	IF stCmdModesStates.stStates.Active THEN
		stCmdModesStates.stStates.Active := FALSE;
		gpCh[nChanIdx]^.channel_mc_control.mode_and_state.command_w.to_mode := HLI_IMCM_AUTOMATIC_MODE;
		gpCh[nChanIdx]^.channel_mc_control.mode_and_state.command_w.to_state := HLI_IMCM_PROCESS_ACTIVE;		
		pString := ADR(gpCh[nChanIdx]^.channel_mc_control.mode_and_state.command_w.parameter);			
		pString^ := ProgramName;				
		gpCh[nChanIdx]^.channel_mc_control.mode_and_state.command_semaphor_rw  := TRUE;		
	END_IF
	
	IF stCmdModesStates.stStates.Hold THEN
		stCmdModesStates.stStates.Hold:= FALSE;
		gpCh[nChanIdx]^.channel_mc_control.mode_and_state.command_w.to_mode:= HLI_IMCM_AUTOMATIC_MODE;
		gpCh[nChanIdx]^.channel_mc_control.mode_and_state.command_w.to_state := HLI_IMCM_PROCESS_HOLD;		
		gpCh[nChanIdx]^.channel_mc_control.mode_and_state.command_semaphor_rw  := TRUE;
	END_IF
	
	IF stCmdModesStates.stStates.Reset THEN
		stCmdModesStates.stStates.Reset := FALSE;
		gpCh[nChanIdx]^.channel_mc_control.mode_and_state.command_w.to_mode := HLI_IMCM_AUTOMATIC_MODE;
		gpCh[nChanIdx]^.channel_mc_control.mode_and_state.command_w.to_state:= HLI_IMCM_PROCESS_RESETTING;		
		gpCh[nChanIdx]^.channel_mc_control.mode_and_state.command_semaphor_rw  := TRUE;		
	END_IF
	
	HLI3_ChannelModeAuto := TRUE;
ELSE
	HLI3_ChannelModeAuto := FALSE;
END_IF

END_FUNCTION

// CNC/2 OperationMode/HLI3_ChannelModeManual
FUNCTION HLI3_ChannelModeManual : BOOL
VAR_INPUT	
	nChanIdx: INT;	
END_VAR

VAR_IN_OUT
	stCmdModesStates    : ST_CNCCmdModesStates;	
END_VAR

VAR
	pString: POINTER TO STRING;
END_VAR

(* ========================================================= *)
(*    FUN: HLI_ChannelModeManual                             *)
(* --------------------------------------------------------- *)
(*   Desc: switch channel to Manual mode / xxx               *)
(*   Author: MK, MiB, TV, RCH                                *)
(*   Date: 03.03.2017                                        *)
(*   Rev.: 1.5                                               *)
(* ========================================================= *)

IF (NOT  gpCh[nChanIdx]^.channel_mc_control.mode_and_state.command_semaphor_rw) THEN    (* only if semaphor is FALSE...... *)
	IF stCmdModesStates.stStates.Selected THEN
		stCmdModesStates.stStates.Selected := FALSE;
		gpCh[nChanIdx]^.channel_mc_control.mode_and_state.command_w.to_mode := HLI_IMCM_MANUAL_MODE;
		gpCh[nChanIdx]^.channel_mc_control.mode_and_state.command_w.to_state := HLI_IMCM_PROCESS_SELECTED;		
		pString := ADR(gpCh[nChanIdx]^.channel_mc_control.mode_and_state.command_w.parameter);			
		pString^ := '';	
		gpCh[nChanIdx]^.channel_mc_control.mode_and_state.command_semaphor_rw := TRUE;		
	END_IF
	
	IF stCmdModesStates.stStates.Ready THEN
		stCmdModesStates.stStates.Ready := FALSE;
		gpCh[nChanIdx]^.channel_mc_control.mode_and_state.command_w.to_mode := HLI_IMCM_MANUAL_MODE;
		gpCh[nChanIdx]^.channel_mc_control.mode_and_state.command_w.to_state := HLI_IMCM_PROCESS_READY;		
		pString := ADR(gpCh[nChanIdx]^.channel_mc_control.mode_and_state.command_w.parameter);			
		pString^ := '';
		gpCh[nChanIdx]^.channel_mc_control.mode_and_state.command_semaphor_rw := TRUE;		
	END_IF
	
	IF stCmdModesStates.stStates.Active THEN
		stCmdModesStates.stStates.Active := FALSE;
		gpCh[nChanIdx]^.channel_mc_control.mode_and_state.command_w.to_mode := HLI_IMCM_MANUAL_MODE;
		gpCh[nChanIdx]^.channel_mc_control.mode_and_state.command_w.to_state := HLI_IMCM_PROCESS_ACTIVE;		
		pString := ADR(gpCh[nChanIdx]^.channel_mc_control.mode_and_state.command_w.parameter);			
		pString^ := '';						
		gpCh[nChanIdx]^.channel_mc_control.mode_and_state.command_semaphor_rw := TRUE;	
	END_IF
	
	IF stCmdModesStates.stStates.Hold THEN
		stCmdModesStates.stStates.Hold := FALSE;
		gpCh[nChanIdx]^.channel_mc_control.mode_and_state.command_w.to_mode := HLI_IMCM_MANUAL_MODE;
		gpCh[nChanIdx]^.channel_mc_control.mode_and_state.command_w.to_state := HLI_IMCM_PROCESS_HOLD;		
		gpCh[nChanIdx]^.channel_mc_control.mode_and_state.command_semaphor_rw := TRUE;		
	END_IF
	
	IF stCmdModesStates.stStates.Reset THEN
		stCmdModesStates.stStates.Reset := FALSE;
		gpCh[nChanIdx]^.channel_mc_control.mode_and_state.command_w.to_mode:= HLI_IMCM_MANUAL_MODE;
		gpCh[nChanIdx]^.channel_mc_control.mode_and_state.command_w.to_state := HLI_IMCM_PROCESS_RESETTING;		
		gpCh[nChanIdx]^.channel_mc_control.mode_and_state.command_semaphor_rw:= TRUE;		
	END_IF

	HLI3_ChannelModeManual := TRUE;
ELSE
	HLI3_ChannelModeManual := FALSE;
END_IF

END_FUNCTION

// CNC/2 OperationMode/HLI3_ChannelModeMDI
FUNCTION HLI3_ChannelModeMDI : BOOL
VAR_INPUT	
	nChanIdx: INT;	
	/// pointer to the MDI program string 
	pMDIString: POINTER TO STRING(HLI_IMCM_MODE_STATE_PARAM_STRL);
END_VAR

VAR_IN_OUT
	stCmdModesStates    : ST_CNCCmdModesStates;	
END_VAR
VAR
	pString: POINTER TO STRING(HLI_IMCM_MODE_STATE_PARAM_STRL);
END_VAR

(* ========================================================= *)
(*    FUN: HLI_ChannelModeMDI                                *)
(* --------------------------------------------------------- *)
(*   Desc: switch channel to MDI mode / xxx                  *)
(*   Author: MK, TV, MiB, Rch                                *)
(*   Date: 18.07.2002                                        *)
(*   Last: 03.03.2017                      				     *)
(*   Rev.: 1.7                                               *)
(* ========================================================= *)

IF (NOT gpCh[nChanIdx]^.channel_mc_control.mode_and_state.command_semaphor_rw) THEN  (* only if semaphor is FALSE...... *)

	IF stCmdModesStates.stStates.Selected THEN
		stCmdModesStates.stStates.Selected := FALSE;
		gpCh[nChanIdx]^.channel_mc_control.mode_and_state.command_w.to_mode := HLI_IMCM_MDI_MODE;
		gpCh[nChanIdx]^.channel_mc_control.mode_and_state.command_w.to_state := HLI_IMCM_PROCESS_SELECTED;
		pString := ADR(gpCh[nChanIdx]^.channel_mc_control.mode_and_state.command_w.parameter);					
		pString^ := pMDIString^;
		gpCh[nChanIdx]^.channel_mc_control.mode_and_state.command_semaphor_rw := TRUE;		
	END_IF
	
	IF stCmdModesStates.stStates.Ready THEN
		stCmdModesStates.stStates.Ready := FALSE;
		gpCh[nChanIdx]^.channel_mc_control.mode_and_state.command_w.to_mode:= HLI_IMCM_MDI_MODE;
		gpCh[nChanIdx]^.channel_mc_control.mode_and_state.command_w.to_state := HLI_IMCM_PROCESS_READY;		
		gpCh[nChanIdx]^.channel_mc_control.mode_and_state.command_semaphor_rw := TRUE;		
	END_IF
	
	IF stCmdModesStates.stStates.Active THEN
		stCmdModesStates.stStates.Active := FALSE;
		gpCh[nChanIdx]^.channel_mc_control.mode_and_state.command_w.to_mode := HLI_IMCM_MDI_MODE;
		gpCh[nChanIdx]^.channel_mc_control.mode_and_state.command_w.to_state := HLI_IMCM_PROCESS_ACTIVE;
		pString := ADR(gpCh[nChanIdx]^.channel_mc_control.mode_and_state.command_w.parameter);					
		pString^ := pMDIString^;
		gpCh[nChanIdx]^.channel_mc_control.mode_and_state.command_semaphor_rw := TRUE;		
	END_IF
	
	IF stCmdModesStates.stStates.Hold THEN
		stCmdModesStates.stStates.Hold := FALSE;
		gpCh[nChanIdx]^.channel_mc_control.mode_and_state.command_w.to_mode := HLI_IMCM_MDI_MODE;
		gpCh[nChanIdx]^.channel_mc_control.mode_and_state.command_w.to_state:= HLI_IMCM_PROCESS_HOLD;		
		gpCh[nChanIdx]^.channel_mc_control.mode_and_state.command_semaphor_rw := TRUE;		
	END_IF
	
	IF stCmdModesStates.stStates.Reset THEN
		stCmdModesStates.stStates.Reset := FALSE;
		gpCh[nChanIdx]^.channel_mc_control.mode_and_state.command_w.to_mode := HLI_IMCM_MDI_MODE;
		gpCh[nChanIdx]^.channel_mc_control.mode_and_state.command_w.to_state := HLI_IMCM_PROCESS_RESETTING;		
		gpCh[nChanIdx]^.channel_mc_control.mode_and_state.command_semaphor_rw := TRUE;		
	END_IF
	HLI3_ChannelModeMDI := TRUE;	
ELSE
	HLI3_ChannelModeMDI := FALSE;
END_IF

END_FUNCTION

// CNC/2 OperationMode/HLI3_ChannelModeReference
FUNCTION HLI3_ChannelModeReference : BOOL
VAR_INPUT	
	nChanIdx: INT;	
	/// the referencing string 
	sRefPosString: STRING(HLI_IMCM_MODE_STATE_PARAM_STRL);	
END_VAR

VAR_IN_OUT
	stCmdModesStates    : ST_CNCCmdModesStates;	
END_VAR

VAR
	pString: POINTER TO STRING(HLI_IMCM_MODE_STATE_PARAM_STRL);
END_VAR

(* ========================================================= *)
(*    FUN: HLI_ChannelModeReference                          *)
(* --------------------------------------------------------- *)
(*   Desc: switch channel to Reference mode / xxx            *)
(*   Author: MK, MiB, TV                                     *)
(*   Date: 03.03.2017                                        *)
(*   Rev.: 1.5                                               *)
(* ========================================================= *)


(************************************************************
	RefPosString:
	Element: parameter ( ASCII char set, Länge:256 Zeichen)

	Vorgabe zur Parametrierung der Referenzpunktfahrt.

	Ist dieser STRING leer, so wird defaultmäßig das
	Automatikprogramm "rpf.nc" angewählt.

	Ansonsten kann durch explizite Angabe der Achsen und
	Zeitpunkt im Format "G74
	<Achsbezeichner_1><Zeitpunkt_1> ...
	<Achsbezeichner_n><Zeitpunkt_n>"
	eine individuelle Referenzpunktfahrt vorgegeben werden.
*************************************************************)

IF (NOT gpCh[nChanIdx]^.channel_mc_control.mode_and_state.command_semaphor_rw) THEN  (* only if semaphor is FALSE...... *)
	IF stCmdModesStates.stStates.Selected THEN
		stCmdModesStates.stStates.Selected := FALSE;
		gpCh[nChanIdx]^.channel_mc_control.mode_and_state.command_w.to_mode := HLI_IMCM_REFERENCE_MODE;
		gpCh[nChanIdx]^.channel_mc_control.mode_and_state.command_w.to_state := HLI_IMCM_PROCESS_SELECTED;		
		gpCh[nChanIdx]^.channel_mc_control.mode_and_state.command_semaphor_rw := TRUE;	
	END_IF
	
	IF stCmdModesStates.stStates.Ready THEN
		stCmdModesStates.stStates.Ready := FALSE;
		gpCh[nChanIdx]^.channel_mc_control.mode_and_state.command_w.to_mode := HLI_IMCM_REFERENCE_MODE;
		gpCh[nChanIdx]^.channel_mc_control.mode_and_state.command_w.to_state := HLI_IMCM_PROCESS_READY;		
		pString := ADR(gpCh[nChanIdx]^.channel_mc_control.mode_and_state.command_w.parameter);	
		gpCh[nChanIdx]^.channel_mc_control.mode_and_state.command_semaphor_rw := TRUE;		
	END_IF
	
	IF stCmdModesStates.stStates.Active THEN
		stCmdModesStates.stStates.Active := FALSE;
		gpCh[nChanIdx]^.channel_mc_control.mode_and_state.command_w.to_mode := HLI_IMCM_REFERENCE_MODE;
		gpCh[nChanIdx]^.channel_mc_control.mode_and_state.command_w.to_state := HLI_IMCM_PROCESS_ACTIVE;		
		pString := ADR(gpCh[nChanIdx]^.channel_mc_control.mode_and_state.command_w.parameter);	
		pString^ := sRefPosString;
		gpCh[nChanIdx]^.channel_mc_control.mode_and_state.command_semaphor_rw:= TRUE;		
	END_IF
	
	IF stCmdModesStates.stStates.Hold THEN
		stCmdModesStates.stStates.Hold := FALSE;
		gpCh[nChanIdx]^.channel_mc_control.mode_and_state.command_w.to_mode := HLI_IMCM_REFERENCE_MODE;
		gpCh[nChanIdx]^.channel_mc_control.mode_and_state.command_w.to_state := HLI_IMCM_PROCESS_HOLD;		
		gpCh[nChanIdx]^.channel_mc_control.mode_and_state.command_semaphor_rw := TRUE;		
	END_IF
	
	IF stCmdModesStates.stStates.Reset THEN
		stCmdModesStates.stStates.Reset := FALSE;
		gpCh[nChanIdx]^.channel_mc_control.mode_and_state.command_w.to_mode:= HLI_IMCM_REFERENCE_MODE;
		gpCh[nChanIdx]^.channel_mc_control.mode_and_state.command_w.to_state := HLI_IMCM_PROCESS_RESETTING;		
		gpCh[nChanIdx]^.channel_mc_control.mode_and_state.command_semaphor_rw := TRUE;		
	END_IF

	HLI3_ChannelModeReference := TRUE;
ELSE
	HLI3_ChannelModeReference := FALSE;
END_IF

END_FUNCTION

// CNC/2 OperationMode/HLI3_ChannelModeStandby
FUNCTION HLI3_ChannelModeStandby : BOOL
VAR_INPUT	 
	nChanIdx: INT;
	ProgramName: STRING(HLI_IMCM_MODE_STATE_PARAM_STRL);			
END_VAR

VAR_IN_OUT
	stCmdModesStates    : ST_CNCCmdModesStates;	
END_VAR

VAR
	pString: POINTER TO STRING(HLI_IMCM_MODE_STATE_PARAM_STRL);
	nCHan: INT;
END_VAR

(* ========================================================= *)
(*    FUN: HLI_ChannelModeStandby                            *)
(* --------------------------------------------------------- *)
(*   Desc: switch channel to Standby mode / xxx              *)
(*   Author: MK, MiB, TV                                     *)
(*   Date: 16.05.2018                                        *)
(*   Rev.: 1.6                                               *)
(* ========================================================= *)

IF (NOT gpCh[nChanIdx]^.channel_mc_control.mode_and_state.command_semaphor_rw) THEN  (* only if semaphor is FALSE...... *)
	IF stCmdModesStates.stStates.Selected THEN
		stCmdModesStates.stStates.Selected := FALSE;
		gpCh[nChanIdx]^.channel_mc_control.mode_and_state.command_w.to_mode := HLI_IMCM_STANDBY_MODE;
		gpCh[nChanIdx]^.channel_mc_control.mode_and_state.command_w.to_state := HLI_IMCM_PROCESS_SELECTED;
		pString := ADR(gpCh[nChanIdx]^.channel_mc_control.mode_and_state.command_w.parameter);			
		pString^ := ProgramName;				
		gpCh[nChanIdx]^.channel_mc_control.mode_and_state.command_semaphor_rw := TRUE;		
	END_IF
	
	IF stCmdModesStates.stStates.Ready THEN
		stCmdModesStates.stStates.Ready := FALSE;
		gpCh[nChanIdx]^.channel_mc_control.mode_and_state.command_w.to_mode := HLI_IMCM_STANDBY_MODE;
		gpCh[nChanIdx]^.channel_mc_control.mode_and_state.command_w.to_state := HLI_IMCM_PROCESS_READY;		
		pString := ADR(gpCh[nChanIdx]^.channel_mc_control.mode_and_state.command_w.parameter);			
		pString^ := ProgramName;	
		gpCh[nChanIdx]^.channel_mc_control.mode_and_state.command_semaphor_rw := TRUE;		
	END_IF
	
	IF stCmdModesStates.stStates.Active THEN
		stCmdModesStates.stStates.Active := FALSE;
		gpCh[nChanIdx]^.channel_mc_control.mode_and_state.command_w.to_mode := HLI_IMCM_STANDBY_MODE;
		gpCh[nChanIdx]^.channel_mc_control.mode_and_state.command_w.to_state := HLI_IMCM_PROCESS_ACTIVE;		
		pString := ADR(gpCh[nChanIdx]^.channel_mc_control.mode_and_state.command_w.parameter);			
		pString^ := ProgramName;	
		gpCh[nChanIdx]^.channel_mc_control.mode_and_state.command_semaphor_rw := TRUE;		
	END_IF
	
	IF stCmdModesStates.stStates.Hold THEN
		stCmdModesStates.stStates.Hold := FALSE;
		gpCh[nChanIdx]^.channel_mc_control.mode_and_state.command_w.to_mode := HLI_IMCM_STANDBY_MODE;
		gpCh[nChanIdx]^.channel_mc_control.mode_and_state.command_w.to_state:= HLI_IMCM_PROCESS_HOLD;		
		gpCh[nChanIdx]^.channel_mc_control.mode_and_state.command_semaphor_rw := TRUE;	
	END_IF
	
	IF stCmdModesStates.stStates.Reset THEN
		stCmdModesStates.stStates.Reset := FALSE;
		gpCh[nChanIdx]^.channel_mc_control.mode_and_state.command_w.to_mode := HLI_IMCM_STANDBY_MODE;
		gpCh[nChanIdx]^.channel_mc_control.mode_and_state.command_w.to_state:= HLI_IMCM_PROCESS_RESETTING;		
		gpCh[nChanIdx]^.channel_mc_control.mode_and_state.command_semaphor_rw := TRUE;		
	END_IF
	
	HLI3_ChannelModeStandby := TRUE;
ELSE
	HLI3_ChannelModeStandby := FALSE;
END_IF

END_FUNCTION

// CNC/2 OperationMode/HLI3_ChannelReset
FUNCTION HLI3_ChannelReset : BOOL
VAR_INPUT
	/// Channel index 
	nChanIdx: INT;
END_VAR
VAR
	/// local pointer to Data of actual Channel 
	pChannelData: POINTER TO HIGH_LEVEL_INTERFACE_CH;
END_VAR

(* ========================================================= 	*)
(*    FUN: HLI_ChannelReset                                  	*)
(* --------------------------------------------------------- 	*)
(*   Desc:                                                   	*)
(* 	 Author: MK ,MiB, TV                                       	*)
(*   Date: 17.01.2018                                        	*)
(*   Rev.: 1.3                                               	*)
(* 	1.2 16.04.2019 Set and Reset the flag  bStateResetting in 	*)
(* 	CNCSystem structur											*)
(*  1.3 31.01.2022 Reset tool request on resetting				*)
(* ========================================================= 	*)

HLI3_ChannelReset := FALSE;
IF NOT HLI3_CheckChannelValid(nChannel := nChanIdx) THEN
	RETURN;
END_IF

(* get pointer to channel data *)
pChannelData := gpCh[nChanIdx];
IF (pChannelData = 0) THEN   (* check for zero pointer *)
	RETURN;
END_IF


CNCSystem.Channel[nChanIdx].bStateResetting := FALSE;

(* is a reset commanded *)
IF pChannelData^.bahn_lc_control.plc_reset.command_r = TRUE THEN
	
	CNCSystem.Channel[nChanIdx].bStateResetting := TRUE;

	(* Reset all M- and H-Functions whenn the channel gets resetted *)
	HLI3_ChannelResetMFunctions(nChanIdx);
	HLI3_ChannelResetHFunctions(nChanIdx);
	
	(* Reset tool request *)
	CNCSystem.Channel[nChanIdx].ToolData.bOldToolDataExist := FALSE;
	CNCSystem.Channel[nChanIdx].ToolData.bToolRequest := FALSE;
	CNCSystem.Channel[nChanIdx].ToolData.bResetToolRequest := TRUE;
	CNCSystem.Channel[nChanIdx].ToolDataJson.bResetToolRequest := TRUE;			
	
	(* quit this reset *)
	pChannelData^.bahn_lc_control.plc_reset.state_w := TRUE;	
	HLI3_ChannelReset := TRUE;
END_IF

END_FUNCTION

// CNC/4 MHT-Function/HLI3_ChannelResetMFunctions
FUNCTION HLI3_ChannelResetMFunctions : BOOL
VAR_INPUT
	/// Channel number 
	nChanIdx: INT;
END_VAR
VAR
	idx: INT;
END_VAR

(* ========================================================= *)
(*    FUN: HLI_ChannelResetMFunctions                        *)
(* --------------------------------------------------------- *)
(*   Desc:                                                   *)
(* Author: MK                                                *)
(*   Date: 10.05.2007                                        *)
(*   Rev.: 1.00                                              *)
(*         1.1   Reset starts at M0 insteat of M1            *)
(* ========================================================= *)

IF NOT HLI3_CheckChannelValid(nChannel := nChanIdx) THEN
	HLI3_ChannelResetMFunctions := FALSE;
	RETURN; (* A b b r u c h *)
END_IF


FOR idx := 0 TO 999 DO
	CNCSystem.Channel[nChanIdx].M[idx].bState_rw := FALSE;
	CNCSystem.Channel[nChanIdx].M[idx].bRes := FALSE;
	CNCSystem.Channel[nChanIdx].actM_r :='';
END_FOR

HLI3_ChannelResetMFunctions := TRUE;

END_FUNCTION

// CNC/4 MHT-Function/HLI3_ChannelResetHFunctions
FUNCTION HLI3_ChannelResetHFunctions : BOOL
VAR_INPUT
	/// Channel number 
	nChanIdx: INT;
END_VAR
VAR
	idx: INT;
END_VAR

(* ========================================================= *)
(*    FUN: HLI_ChannelResetHFunctions                        *)
(* --------------------------------------------------------- *)
(*   Desc:                                                   *)
(* Author: MiB                                                *)
(*   Date: 23.11.2012                                        *)
(*   Rev.: 1.1                                              *)
(* ========================================================= *)



IF NOT HLI3_CheckChannelValid(nChannel := nChanIdx) THEN
	HLI3_ChannelResetHFunctions := FALSE;
	RETURN; (* A b b r u c h *)
END_IF


FOR idx := 0 TO 999 DO
	CNCSystem.Channel[nChanIdx].H[idx].bState_rw := FALSE;
	CNCSystem.Channel[nChanIdx].H[idx].bRes := FALSE;
	CNCSystem.Channel[nChanIdx].actH_r :='';
END_FOR

HLI3_ChannelResetHFunctions := TRUE;

END_FUNCTION

// CNC/2 OperationMode/HLI3_ChannelResetRequest
FUNCTION_BLOCK HLI3_ChannelResetRequest
VAR_INPUT
	bExec: BOOL;
	/// Channel number 
	nChanIdx: INT;
	pChannel: POINTER TO ST_CncChannel;
END_VAR
VAR_OUTPUT
	bBusy: BOOL;
	bSwitchMode: BOOL;
	nMode: UDINT;
END_VAR
VAR
	fbRtrigExec: R_TRIG;
	/// Index of channel specific HLI area 
	nHliChIfcIdx: INT;
	nState: UINT;
	pCommand: POINTER TO HLI_PROC_TRANS_TO_MODE_STATE;
	actualMode: UDINT;
	fbTON: TON;
END_VAR

(******************************************************************************)
(* POU:				HLI_ChannelResetRequest									*)
(* Type:				Function block										*)
(* Customer:		Common													*)
(* Date:				07/11/16											*)
(* Last:				10/03/10											*)
(* -------------------------------------------------------------------------- *)
(* Revision:		1.0														*)
(* Author:			MiB														*)
(* Description: 	Performs a reset in the given cnc channel. 				*)
(* -------------------------------------------------------------------------- *)
(* Revision:		1.10													*)
(* Author:			MiB														*)
(* Description: 	Changed from PRG to FB.									*)
(* -------------------------------------------------------------------------- *)
(* Revision:		2.00															*)
(* Author:			HR																*)
(* Description: 	Deleted references to global variable 'PLCMachineMode[n]'.		*)
(*						The FB now works with VAR_OUTPUT 'nMode' and 'bSwitchMode'	*)
(*						as a callback to the initiator to let it perform the change	*)
(*						of the operation mode by itself in order to reset the cnc	*)
(*						channel.													*)
(* -------------------------------------------------------------------------- *)
(* Revision:		2.01																			*)
(* Author:			TV																				*)
(* Description: 	Expand State "Wait for previous mode"  *)
(*				Prevent to trigger the state machine during the mode switch							*)
(* -------------------------------------------------------------------------- *)
(* Revision:		2.02																			*)
(* Author:			MiB																				*)
(* Description: 	Tc3*)
(******************************************************************************)


fbRtrigExec( clk := bExec   );

IF fbRtrigExec.Q THEN
	bBusy := TRUE;
	nState := 10;
END_IF


CASE nState OF

0:		(* IDLE *)
		bBusy := FALSE;

10:	(* Reset request: get actual opmode *)
		bSwitchMode := FALSE;
		actualMode := gpCh[nChanIdx]^.channel_mc_control.mode_and_state.state_r.mode;
		nState := nState + 10;

20:  (* switch to standby *)
		bSwitchMode := TRUE;
		nMode:= HLI_IMCM_STANDBY_MODE;
		fbTON(IN:= FALSE);
		nState := nState + 10;

30: 	(* Wait for modeswitch *)
		bSwitchMode := FALSE;
		fbTON(IN:= TRUE, PT:= t#2000ms);
	 	IF gpCh[nChanIdx]^.channel_mc_control.mode_and_state.state_r.mode = HLI_IMCM_STANDBY_MODE THEN
			nState := nState + 10;
		END_IF
		IF fbTON.Q THEN
			(* Timeout Error -> go on with next step *)
			nState := nState + 10;
		END_IF

40:	(* switch back to previous mode *)
		bSwitchMode := TRUE;
		nMode:= actualMode;
		fbTON(IN:= FALSE);
		nState := nState + 10;

50:	(* Wait for previous mode  *)
		fbTON(IN:= TRUE, PT:= t#2000ms);
		IF (gpCh[nChanIdx]^.channel_mc_control.mode_and_state.state_r.mode = 	actualMode) THEN
			nState := nState + 10;
		END_IF
		IF fbTON.Q THEN
			(* Timeout Error -> go on with next step *)
			nState := nState + 10;
		END_IF

60: 	(* ready *)
		bSwitchMode := FALSE;
		nState := 0;

END_CASE



(* das muss ins aufrufende Programm: (HLI_CNCChannel)

VAR
	bResetRequest:			BOOL;
	fbRTrigReset:			R_TRIG;
	ChannelResetRequest: HLI_ChannelResetRequest;
END_VAR

fbRTrigReset(clk := bStateReset);
IF fbRTrigReset.Q THEN
	bResetRequest := TRUE;
	...
END_IF

(* Handle Channel reset *)
ChannelResetRequest
	(bExec 		:= bResetRequest ,
	 nChan 		:= nChan,
	 pChannel	:= ADR(CNCSystem.Channel[nChan])
	);

IF ChannelResetRequest.bSwitchMode THEN
	bModeStandby	:= bModeStandby OR (ChannelResetRequest.nMode = HLI_IMCM_STANDBY_MODE);
	bModeAutomatic	:= bModeAutomatic OR (ChannelResetRequest.nMode = HLI_IMCM_AUTOMATIC_MODE);
	bModeManual		:= bModeManual OR (ChannelResetRequest.nMode = HLI_IMCM_MANUAL_MODE);
	bModeMDI			:= bModeMDI OR (ChannelResetRequest.nMode = HLI_IMCM_MDI_MODE);
	bModeReference	:= bModeReference OR (ChannelResetRequest.nMode = HLI_IMCM_REFERENCE_MODE);
END_IF

IF bResetRequest AND NOT ChannelResetRequest.bBusy THEN
	bResetRequest := FALSE;
END_IF

*)

END_FUNCTION_BLOCK

// CNC/2 OperationMode/HLI3_CNCChannel
FUNCTION_BLOCK HLI3_CNCChannel
VAR_INPUT
	/// index of channel
	nChanIdx: INT;
 
	bCmdAutomatic : BOOL;
	bCmdManual : BOOL;
    bCmdReference : BOOL;
    bCmdMDI : BOOL;		
	bCmdStandby: BOOL;
	bCmdStart : BOOL;
	bCmdStop  : BOOL;
	bCmdReset : BOOL;		
	/// must be xxx.nc 
	sProgramName: STRING(HLI_IMCM_MODE_STATE_PARAM_STRL);
	/// the MDI string 
	sMDIString: STRING(HLI_IMCM_MODE_STATE_PARAM_STRL);
	/// static signal 
	bBackwardMotion: BOOL;
	/// static signal 
	bFeedHold: BOOL;
	/// static signal 
	bReducedFeed: BOOL;
	/// static signal 
	bSingleBlock: BOOL;
	/// static signal 
	bPrgBlockIgnore: BOOL;
	/// static signal 
	bM01Stop: BOOL;
	/// static signal 
	nSyntaxCheck: DINT;		
	// Manual Mode
	stManualModeParameter: ST_ManualModeParameter;
	stManualModeControlElements: ST_ManualModeControlElements;
	// M30 Acknowledgement inside Channel FB
	bM30Acknowledgement : BOOL;
	// Override 
	nFeedOverride : UINT;
	nRapidFeedOverride : UINT;
	bEmergencyStop : BOOL;
	stOptions : ST_CNC_CH_Options;
END_VAR

VAR_OUTPUT
	bError 	: BOOL;	
	nErrorID	: UDINT;
END_VAR

VAR_IN_OUT
	/// please only a flank 
	bModeStandby: BOOL;
	/// please only a flank 
	bModeAutomatic: BOOL;
	/// please only a flank 
	bModeManual: BOOL;
	/// please only a flank 
	bModeMDI: BOOL;
	/// please only a flank 
	bModeReference: BOOL;
	/// please only a flank 
	bStateSelect: BOOL;
	/// please only a flank 
	bStateReady: BOOL;
	/// please only a flank 
	bStateStart: BOOL;
	/// please only a flank 
	bStateStop: BOOL;
	/// please only a flank 
	bStateReset: BOOL;
	/// please only a flank 
	bDoSingleBlock: BOOL;
	// manual mode
	stManualModeControlElementState: ST_ManualModeControlElementState;
END_VAR
VAR
	bGoToActive	: BOOL;	 	
	/// Pointer to channel control structure 
	pChannel: POINTER TO ST_CncChannel;
	ChannelMHTFunction: HLI3_QuitChannelMHTFunction;
	/// Current Mode of Operation Modes;
	currentMode: UDINT;
	/// Current State of Operation Modes;
	currentState: UDINT;
	idx: INT;	
	bCheckOpModeFirst: BOOL;
	fbRTrigReset: R_TRIG;
	bResetRequest: BOOL;	
	nStateAutoMDIStart: INT;
	ModeManual : HLI3_ManualModeHandler;	
	fbToolDataJson: FB_ToolDataJson;
	stCmdModesStates    : ST_CNCCmdModesStates;

	fbRTrigCmdStart: R_TRIG;
	fbRTrigCmdStop:  R_TRIG;
	fbRTrigCmdReset: R_TRIG;	
	fbRTrigCmdAutomatic : R_TRIG;
	fbRTrigCmdManual : R_TRIG;
    fbRTrigCmdReference : R_TRIG;
    fbRTrigCmdMDI : R_TRIG;		
	fbRTrigCmdStandby: R_TRIG;
	// File Offset
	fbADSWrite : ADSWRITE;	  
	fbRTrigSetFileOffset: R_TRIG;	
	nState : INT;	
END_VAR

(* ========================================================= *)
(*     FB: HLI_CNCChannel                                    *)
(* --------------------------------------------------------- *)
(*   Desc:                                                   *)
(*   Author: MK ,MiB, TV, Rch                                *)
(*   Date: 2020.07.27                                        *)
(*   Rev.: 1.21                                              *)
(*         1.2 Before "start" the state is swicthed to 		 *)
(*				"Selected" and "Ready" to ensure that the    *)	
(*				actual selected program will start 			 *)
(*		   	1.3  BugFix : nChanNo at HLI3_ChannelModeMDI()    *)
(*         	1.4  Implement state switch to "selected" and "ready"  *)         
(*		   	1.5  Channel reset via commanding state 			 *)
(*              RESETTING directly							 *)  
(*		   	1.6  Optimized Channel reset via commanding state *)
(*				RESETTING directly						     *)
(*		   	1.7  Init Paramerer for Manual mode as input parameter*)
(*		   	1.8  BugFix : max index for HLI3_AxisReset		*)
(*		   	1.9  Implementation of HLI3_ManualModeHandler	*)
(*		   	1.10 Implementation of Input bM30Acknowledgement	*)
(*		   	1.12 Optimized Operating modes					*)
(*		   	1.13 Optimized Operating modes				    *)
(*		   	1.14 Optimized M and H Function during Reset     *)
(*		   	1.15 Implementation of ST_CNC_CH_Options Structure *)
(*		   	1.16 BugFix: bCmdReset in mode "Standby" now working *)
(*			1.17 Implementation of CNC PLC Watchdog			*)  
(*			1.18 Optimized CNC PLC Watchdog					*)
(*			1.18 Optimized G201 ManualMode					*)
(*			1.19 Add CmdStandby 							*)
(*			1.20 New Manual Mode 							*)
(*			1.21 Option bDisableAutoAcknowledgeM 			*)
(*			1.22 Option program start with file Offset 		*)
(*          1.23 use FB_ToolDataJson if enabled in global Variable CNCSystem.bToolDataJson *)
(* =========================================================*)

IF NOT HLI3_CheckChannelValid(nChannel := nChanIdx) THEN
	RETURN;
END_IF

// CNC PLC Watchdog	
IF NOT stOptions.bDisableCNCPLCWatchDog THEN
	HLI3_SetPLCAlive(nChanIdx :=  nChanIdx);
END_IF

(* handle reset request *)
fbRTrigReset
	(CLK := bStateReset);
	
IF fbRTrigReset.Q THEN
	nStateAutoMDIStart := 0;
END_IF

// FileOffset
FileOffset();

fbRTrigCmdAutomatic(CLK:=bCmdAutomatic);
fbRTrigCmdManual(CLK:=bCmdManual);
fbRTrigCmdReference(CLK:=bCmdReference);
fbRTrigCmdMDI(CLK:=bCmdMDI);
fbRTrigCmdStandby(CLK:=bCmdStandby);	

fbRTrigCmdStart(CLK:=bCmdStart);  
fbRTrigCmdStop(CLK:=bCmdStop);
fbRTrigCmdReset(CLK:=bCmdReset);

(* ************************************* *)
(*  Motion-Control                       *)
(* ************************************* *)

(* EmergencyStop *)
HLI3_ChannelSetEmergencyStop(nChanIdx:=nChanIdx, bEStop := bEmergencyStop);
 
(* Feed Override [0.1%] *)
HLI3_SetChannelOverride(nChanIdx:=nChanIdx, nOverride := nFeedOverride);

(* Rapid feed override [0.1%], must be activated with parameter P-CHAN-00181 *)
HLI3_SetChannelRapidOverride(nChanIdx:=nChanIdx, nOverride := nRapidFeedOverride);

(* Backward Motion *)
HLI3_ChannelSetBackwardMotion(nChanIdx:=nChanIdx, bBackwardMotion:=bBackwardMotion);

(* Program Block Ignore *)
HLI3_ChannelSetProgramBlockIgnore(nChanIdx:=nChanIdx, bPrgBlockIgnore:=bPrgBlockIgnore);

(* Feed Hold *)
HLI3_ChannelSetFeedHold(nChanIdx:=nChanIdx, bFeedHold:=bFeedHold);

(* Single Step *)
HLI3_ChannelSetSingleBlock(nChanIdx:=nChanIdx, bSingleBlock:=bSingleBlock);

(* Reduced Feed *)
HLI3_ChannelSetReducedFeed(nChanIdx:=nChanIdx, bReducedFeed:=bReducedFeed);

(* Syntax Check *)
gpCh[nChanIdx]^.decoder_mc_control.execution_mode.command_w := nSyntaxCheck;

(* Optional stop M01 *)
gpCh[nChanIdx]^.bahn_mc_control.m01_stop_enable.command_w := bM01Stop;

(* ************************************ *)
(*  MHT-Function                        *)
(* ************************************ *)

(* MHT-Function, channel *)
IF NOT stOptions.bDisableMFunctHandling THEN
	ChannelMHTFunction(nChanIdx:=nChanIdx, bM30Acknowledgement := bM30Acknowledgement, bDisableAutoAcknowledgeM := stOptions.bDisableAutoAcknowledgeM);
END_IF

(* ************************************* *)
(*  Channel Status Info and error        *)
(* ************************************* *)
HLI3_GetChannelStatusInfo(nChanIdx:=nChanIdx);
HLI3_GetChannelError(nChanIdx:=nChanIdx);

(* ************************************* *)
(*  do single stepping                   *)
(* ************************************* *)
(* Achtung: hier noch anpassen, nur in Abhaengigkeit vom aktuellen Status den Start setzen *)
IF bDoSingleBlock THEN
	bDoSingleBlock := FALSE;
	bStateStart 	:= TRUE;
END_IF

(* ************************************* *)
(*  Operation Modes                      *)
(* ************************************* *)
(* Target modes and states *)
pChannel := ADR(CNCSystem.Channel[nChanIdx]);
OpModes();

(* OperationMode Standby *)
IF stCmdModesStates.stModes.Standby = TRUE THEN
	HLI3_ChannelModeStandby(nChanIdx := nChanIdx,ProgramName:=sProgramName, stCmdModesStates:=stCmdModesStates);
END_IF

(* OperationMode Auto *)
IF stCmdModesStates.stModes.Auto = TRUE THEN
	HLI3_ChannelModeAuto(nChanIdx := nChanIdx, ProgramName:=sProgramName, stCmdModesStates:=stCmdModesStates );
END_IF

(* OperationMode MDI *)
IF stCmdModesStates.stModes.MDI THEN
	(*sProgramName := PLCCncMDIString;*)
	HLI3_ChannelModeMDI(nChanIdx := nChanIdx, pMDIString:=ADR(sMDIString),stCmdModesStates:=stCmdModesStates);
END_IF

(* OperationMode Reference *)
IF stCmdModesStates.stModes.Homing THEN
	sProgramName := '';	(* we choose the default program: rpf.nc *)
	HLI3_ChannelModeReference(nChanIdx := nChanIdx, sRefPosString:=sProgramName, stCmdModesStates:=stCmdModesStates);
END_IF

(* OperationMode Manual *)
(*
IF stCmdModesStates.stModes.Manual THEN	
	HLI3_ChannelModeManual(nChanIdx := nChanIdx, stCmdModesStates:=stCmdModesStates);
END_IF
*)

ModeManual
	(stManualModeParameter  	 	 := stManualModeParameter,
	 stManualModeControlElements	 := stManualModeControlElements,
	 stManualModeControlElementState := stManualModeControlElementState,
	 stCmdModesStates				 := stCmdModesStates,  	
	 arrAxisInG201 				      => stManualModeState[nChanIdx].arrAxisInG201
);
			
IF CNCSystem.bToolDataJson THEN   // tool data transfer via json is enabled
	fbToolDataJson(nChanIdx := nChanIdx);
END_IF


(* Reset *)
HLI3_ChannelReset(nChanIdx:=nChanIdx);							(* channel *)
FOR idx := 0 TO UDINT_TO_INT(gNrAx-1) DO							(* axis *)
	HLI3_AxisReset(nChanNo:=nChanIdx+1, nHliAxisIdx:=idx);
END_FOR

ACTION AutoMDIStart:



CASE nStateAutoMDIStart OF
	0:		;(* IDLE *)
	
	10: (* swicth to selected *)
		stCmdModesStates.stStates.Selected := TRUE;
		nStateAutoMDIStart := nStateAutoMDIStart +10;
		
	20: (* wait for selected *)
		IF (pChannel^.ActState =  HLI_IMCM_PROCESS_SELECTED) THEN
			stCmdModesStates.stStates.Ready := TRUE;
			nStateAutoMDIStart := nStateAutoMDIStart +10;
		END_IF
	30: (* Wait for ready and then start*)
		IF (pChannel^.ActState =  HLI_IMCM_PROCESS_READY) THEN
			stCmdModesStates.stStates.Active := TRUE; 
			nStateAutoMDIStart := 0;
		END_IF
	
END_CASE
END_ACTION

ACTION FileOffset:
fbRTrigSetFileOffset(CLK:=stOptions.bSetCNCProgramFileOffset);
IF fbRTrigSetFileOffset.Q THEN
   	nState 				:= 10;   	   
   	fbADSWrite.WRITE 	:= FALSE;	
	bError				:= FALSE;		
END_IF


CASE nState OF
0:
	;
10: // Write File Offset
	fbADSWrite( NetID := '', Port := 553, IdxGrp := 16#00020100 + INT_TO_UDINT(nChanIdx)+1, IdxOffs := 16#00000011,
         LEN := 4, SrcAddr := ADR(stOptions.nCNCProgramFileOffset), WRITE := TRUE, TMOUT := T#1S);
		 		
	IF NOT fbADSWrite.Busy AND NOT fbADSWrite.Err THEN
			fbADSWrite(WRITE:=FALSE);		
			nState := 0;
		ELSIF NOT fbADSWrite.Busy AND fbADSWrite.Err THEN			
			bError := TRUE;
			nErrorID := fbADSWrite.ERRID; 									
			fbADSWrite(WRITE:=FALSE);
			nState := 0;
		END_IF;
		
		
		
END_CASE
END_ACTION

ACTION OpModes:
(*************************************************)
(* Restore internal state at first run           *)
(* after PLC reset                               *)
(*************************************************)

IF bCheckOpModeFirst = FALSE THEN
	bCheckOpModeFirst := TRUE;
	currentMode := HLI3_GetChannelMode(nChanIdx:=nChanIdx);
	IF currentMode = HLI_IMCM_STANDBY_MODE THEN
		stCmdModesStates.stModes.Standby := TRUE;
	END_IF
	IF currentMode = HLI_IMCM_AUTOMATIC_MODE THEN
		stCmdModesStates.stModes.Auto := TRUE;
	END_IF
	IF currentMode = HLI_IMCM_MDI_MODE THEN
		stCmdModesStates.stModes.MDI := TRUE;
	END_IF
	IF currentMode = HLI_IMCM_MANUAL_MODE THEN
		stCmdModesStates.stModes.Manual := TRUE;
	END_IF
	IF currentMode = HLI_IMCM_REFERENCE_MODE THEN		
		stCmdModesStates.stModes.Homing := TRUE;
	END_IF
END_IF


(*************************************************)
(* Operation Modes                               *)
(*************************************************)

IF bModeStandby OR fbRTrigCmdStandby.Q THEN
	bModeStandby := FALSE;
	stCmdModesStates.stModes.Standby		:= TRUE;
	stCmdModesStates.stModes.Auto			:= FALSE;
	stCmdModesStates.stModes.MDI			:= FALSE;
	stCmdModesStates.stModes.Manual		:= FALSE;
	stCmdModesStates.stModes.Homing		:= FALSE;
	stCmdModesStates.stStates.Selected	:= TRUE;
END_IF

IF bModeAutomatic OR fbRTrigCmdAutomatic.Q THEN
	bModeAutomatic 				:= FALSE;
	bGoToActive					:= FALSE;
	stCmdModesStates.stModes.Standby		:= FALSE;
	stCmdModesStates.stModes.Auto			:= TRUE;
	stCmdModesStates.stModes.MDI			:= FALSE;
	stCmdModesStates.stModes.Manual		:= FALSE;
	stCmdModesStates.stModes.Homing		:= FALSE;

	stCmdModesStates.stStates.Selected	:= TRUE;
END_IF

IF bModeMDI OR fbRTrigCmdMDI.Q THEN
	bModeMDI := FALSE;
	bGoToActive					:= FALSE;
	stCmdModesStates.stModes.Standby		:= FALSE;
	stCmdModesStates.stModes.Auto			:= FALSE;
	stCmdModesStates.stModes.MDI			:= TRUE;
	stCmdModesStates.stModes.Manual		:= FALSE;
	stCmdModesStates.stModes.Homing		:= FALSE;

	stCmdModesStates.stStates.Selected	:= TRUE;
END_IF

IF bModeManual OR fbRTrigCmdManual.Q THEN
	bModeManual := FALSE;
	stCmdModesStates.stModes.Standby		:= FALSE;
	stCmdModesStates.stModes.Auto			:= FALSE;
	stCmdModesStates.stModes.MDI			:= FALSE;
	stCmdModesStates.stModes.Manual		:= TRUE;
	stCmdModesStates.stModes.Homing		:= FALSE;

	stCmdModesStates.stStates.Active		:= TRUE;
END_IF

IF bModeReference OR fbRTrigCmdReference.Q THEN
	bModeReference := FALSE;
	bGoToActive					:= FALSE;
	stCmdModesStates.stModes.Standby		:= FALSE;
	stCmdModesStates.stModes.Auto			:= FALSE;
	stCmdModesStates.stModes.MDI			:= FALSE;
	stCmdModesStates.stModes.Manual		:= FALSE;
	stCmdModesStates.stModes.Homing		:= TRUE;
	
	IF stOptions.bReferenceModeStartRequired THEN
		stCmdModesStates.stStates.Selected	:= TRUE;
	ELSE
		stCmdModesStates.stStates.Active	:= TRUE;			
	END_IF	
	
END_IF



(*************************************************)
(* Operation States                              *)
(*************************************************)

currentMode := HLI3_GetChannelMode(nChanIdx:=nChanIdx);
currentState := HLI3_GetChannelState(nChanIdx:=nChanIdx);

CASE currentMode OF
	(*-------------------------------------------------------------------*)
	HLI_IMCM_STANDBY_MODE:
		IF bStateReset OR fbRTrigCmdReset.Q THEN
			stCmdModesStates.stModes.Standby := TRUE;
			stCmdModesStates.stStates.Reset := TRUE;
		END_IF

	(*-------------------------------------------------------------------*)
	HLI_IMCM_AUTOMATIC_MODE:
		IF bStateStart OR fbRTrigCmdStart.Q THEN  (* replaced a simple 'start' by a sequence which switches the state to selected and ready*)
			IF currentState <> HLI_IMCM_PROCESS_HOLD AND currentState <> HLI_IMCM_PROCESS_ACTIVE THEN
				nStateAutoMDIStart := 10;
			ELSE
				stCmdModesStates.stStates.Active := TRUE; 
			END_IF					   	
		END_IF
		IF nStateAutoMDIStart <> 0 THEN
			AutoMDIStart();
		END_IF

		//IF (bStateStop OR fbRTrigCmdStop.Q) AND currentState <> HLI_IMCM_PROCESS_DESELECTED THEN 
		IF (bStateStop OR fbRTrigCmdStop.Q) AND currentState = HLI_IMCM_PROCESS_ACTIVE THEN           // 2021.05.10 MiB: Stop nur ausführen, wenn gerade "Active" 
			stCmdModesStates.stStates.Hold := TRUE;
		END_IF

		IF bStateReady THEN
			stCmdModesStates.stStates.Ready := TRUE;
		END_IF

		IF bStateReset OR fbRTrigCmdReset.Q THEN
			stCmdModesStates.stStates.Reset := TRUE;
		END_IF
		
		IF bStateSelect THEN
			stCmdModesStates.stStates.Selected := TRUE;
		END_IF		

	(*-------------------------------------------------------------------*)
	HLI_IMCM_MDI_MODE:
		IF bStateStart OR fbRTrigCmdStart.Q THEN
			IF currentState <> HLI_IMCM_PROCESS_HOLD AND currentState <> HLI_IMCM_PROCESS_ACTIVE THEN
				nStateAutoMDIStart := 10;
			ELSE
				stCmdModesStates.stStates.Active := TRUE; 
			END_IF
		END_IF
		
		IF nStateAutoMDIStart <> 0 THEN
			AutoMDIStart();
		END_IF
		
		IF (bStateStop OR fbRTrigCmdStop.Q) AND currentState <> HLI_IMCM_PROCESS_DESELECTED AND currentState = HLI_IMCM_PROCESS_ACTIVE THEN           // 2023.05.24 MiB: only go to "hold" is actstate is active
			stCmdModesStates.stStates.Hold := TRUE;
		END_IF

		IF bStateSelect THEN
			stCmdModesStates.stStates.Selected := TRUE;
		END_IF
		
		IF bStateReady THEN
			stCmdModesStates.stStates.Ready := TRUE;
		END_IF

		IF bStateReset OR fbRTrigCmdReset.Q THEN
			stCmdModesStates.stStates.Reset := TRUE;
		END_IF

	(*-------------------------------------------------------------------*)
	HLI_IMCM_MANUAL_MODE:
		IF bStateStart OR fbRTrigCmdStart.Q OR ((currentState = HLI_IMCM_PROCESS_SELECTED) AND bGoToActive) THEN
			bGoToActive := FALSE;	
			stCmdModesStates.stStates.Active 	:= TRUE;
		END_IF

		IF bStateReady THEN
			stCmdModesStates.stStates.Ready 	:= TRUE;
		END_IF

		IF bStateSelect THEN
			stCmdModesStates.stStates.Selected := TRUE;
		END_IF

		IF bStateStop OR fbRTrigCmdStop.Q THEN
			stCmdModesStates.stStates.Hold := TRUE;
		END_IF

		IF (bStateReset OR fbRTrigCmdReset.Q) THEN	
			stCmdModesStates.stStates.Reset := TRUE;
			IF stCmdModesStates.stModes.Manual THEN
				bGoToActive := TRUE;
			END_IF
		END_IF

	(*-------------------------------------------------------------------*)
	HLI_IMCM_REFERENCE_MODE:
		IF bStateStart OR fbRTrigCmdStart.Q THEN
			stCmdModesStates.stStates.Active := TRUE;
		END_IF

		IF bStateStop OR fbRTrigCmdStop.Q THEN
			stCmdModesStates.stStates.Hold := TRUE;
		END_IF

		IF bStateReset OR fbRTrigCmdReset.Q THEN
			stCmdModesStates.stStates.Reset := TRUE;
		END_IF
END_CASE


bStateStart 	:= FALSE;
bStateStop 		:= FALSE;
bStateReset 	:= FALSE;
bStateSelect 	:= FALSE;
bStateready 	:= FALSE;
END_ACTION

END_FUNCTION_BLOCK

// CNC/7 ToolManagement/FB_ToolDataJson
FUNCTION_BLOCK FB_ToolDataJson
VAR_INPUT
	nChanIdx:   INT;
END_VAR
VAR_OUTPUT
END_VAR
VAR
	nStateTr: INT;
	nStateTrPrep : INT;
	fbJsonParser : FB_JsonDomParser;		
	fbJsonWriter  : FB_JsonSaxWriter;    
 	fbJsonDataType: FB_JsonReadWriteDataType;		
// 	sDataType: STRING;		
	nStateOt : INT;
	nStateEt : INT;	
	sJsonResult : STRING(MAX_JSON_TOOLDATA_SIZE);		
END_VAR

///*********************************************************************************************************
///NAME.......................:		FB_ToolDataJson
///DATUM....................:		27.05.2026
///AUTOR....................:		Michael Balsfulland
///VERSION................:			1.0
///
///Description.: Data transfer of tool data via JSON string to and from ToolDatastructure and HMI				
///**********************************************************************************************************


IF CNCSystem.Channel[nChanIdx].ToolDataJson.bResetToolRequest THEN
	nStateTr := 0;
	nStateTrPrep := 0;
	nStateOt := 0;
	nStateEt := 0;
	sJsonResult := '';
	fbJsonWriter.ResetDocument();
	CNCSystem.Channel[nChanIdx].ToolDataJson.bResetToolRequest := FALSE;	
END_IF


IF CNCSystem.Channel[nChanIdx].ToolData.bToolRequest = true THEN
	IF (nStateTr = 0) THEN     // only if action toolrequest is idle (state == 0)
		nStateTr := 10;
	END_IF
END_IF
a_toolRequest();


IF CNCSystem.Channel[nChanIdx].ToolData.bToolRequestPrepData= TRUE THEN
	IF (nStateTrPrep = 0) THEN     // only if action toolrequest is idle (state == 0)
		nStateTrPrep := 10;
	END_IF
END_IF
b_ToolPrepRequest();


IF CNCSystem.Channel[nChanIdx].ToolData.bOldToolDataExist = TRUE THEN
	IF (nStateOt = 0) THEN
		nStateOt := 10;
	END_IF
END_IF
c_OldToolExists();

IF CNCSystem.Channel[nChanIdx].ToolData.bEditToolDataExist = TRUE THEN
	IF (nStateEt = 0) THEN
		nStateEt := 10;
	END_IF
END_IF
d_EditToolExists();

ACTION a_ToolRequest:




CASE nStateTr OF
	
	10:   // forward request to json DataStructure
		CNCSystem.Channel[nChanIdx].ToolDataJson.nToolRequestID := CNCSystem.Channel[nChanIdx].ToolData.nToolRequestID;
		CNCSystem.Channel[nChanIdx].ToolDataJson.nToolRequestIDSister := CNCSystem.Channel[nChanIdx].ToolData.nToolRequestIDSister;
		CNCSystem.Channel[nChanIdx].ToolDataJson.nToolRequestIDVariant := CNCSystem.Channel[nChanIdx].ToolData.nToolRequestIDVariant;
		CNCSystem.Channel[nChanIdx].ToolDataJson.bToolRequest := TRUE;
		nStateTr := nStateTr + 10;		 		
		
	20:
	   IF CNCSystem.Channel[nChanIdx].ToolDataJson.bToolRequest = FALSE THEN    // wait for received data from HMI   ( bToolRequest is set to false from HMI )
			IF CNCSystem.Channel[nChanIdx].ToolDataJson.PreJsonToToolAcion <> 0 THEN
				nStateTr := nStateTr + 10;    // call the method commit of the ITF
			ELSE 
				nStateTr := nStateTr + 20;	      // go on without ITF
			END_IF	   		   
	   END_IF
	   
	30:
		IF CNCSystem.Channel[nChanIdx].ToolDataJson.PreJsonToToolAcion.Commit(CNCSystem.Channel[nChanIdx].ToolDataJson.stActToolJson) THEN
			CNCSystem.Channel[nChanIdx].ToolDataJson.stActToolJson := CNCSystem.Channel[nChanIdx].ToolDataJson.PreJsonToToolAcion.ToolJson;
			nStateTr := nStateTr + 10;	
		END_IF
	      
	40:	// transfer data from json to plc datastructure		
		IF (SetSymbolFromJson(fbJsonParser.ParseDocument(CNCSystem.Channel[nChanIdx].ToolDataJson.stActToolJson), ADR(CNCSystem.Channel[nChanIdx].ToolData.stActTool))) THEN
			CNCSystem.Channel[nChanIdx].ToolData.bToolRequest := FALSE;
			nStateTr := 0;  // done
		END_IF
				   			   
	
END_CASE
END_ACTION

ACTION b_ToolPrepRequest:

CASE nStateTrPrep OF
	
	10:   // forward request to json DataStructure
		CNCSystem.Channel[nChanIdx].ToolDataJson.nToolRequestPrepId := CNCSystem.Channel[nChanIdx].ToolData.nToolRequestPrepId;
		// Sister and Variant are used if set directly in json request structure, in "old" system sister and variant for prep data was not implemented
		//CNCSystem.Channel[nChanIdx].ToolDataJson.nToolRequestPrepIdSister;
		//CNCSystem.Channel[nChanIdx].ToolDataJson.nToolRequestPrepIdVariant;
		CNCSystem.Channel[nChanIdx].ToolDataJson.bToolRequestPrepData := TRUE;
		nStateTrPrep := nStateTrPrep + 10;		 		
		
	20:
	   IF CNCSystem.Channel[nChanIdx].ToolDataJson.bToolRequestPrepData = FALSE THEN    // wait for received data from HMI   ( bToolRequest is set to false from HMI )
			IF CNCSystem.Channel[nChanIdx].ToolDataJson.PreJsonToToolAcion <> 0 THEN
				nStateTrPrep := nStateTrPrep + 10;    // call the method commit of the ITF
			ELSE 
				nStateTrPrep := nStateTrPrep + 20;	  // go on without ITF
			END_IF	   				   

	   END_IF	

	30:
		IF CNCSystem.Channel[nChanIdx].ToolDataJson.PreJsonToToolAcion.Commit(CNCSystem.Channel[nChanIdx].ToolDataJson.stPrepToolJson) THEN
			CNCSystem.Channel[nChanIdx].ToolDataJson.stPrepToolJson := CNCSystem.Channel[nChanIdx].ToolDataJson.PreJsonToToolAcion.ToolJson;
			nStateTr := nStateTr + 10;	
		END_IF
	      
	40:	
		// transfer data from json to plc datastructure
		IF (SetSymbolFromJson(fbJsonParser.ParseDocument(CNCSystem.Channel[nChanIdx].ToolDataJson.stPrepToolJson), ADR(CNCSystem.Channel[nChanIdx].ToolData.stPrepTool))) THEN
			CNCSystem.Channel[nChanIdx].ToolData.bToolRequestPrepData := FALSE;
			nStateTrPrep := 0;  // done
		END_IF
				   			   
	
END_CASE
END_ACTION

ACTION c_OldToolExists:


CASE nStateOt OF
	
	10:   // forward request to json DataStructure
		  // convert Data to json datastructure
		
		//  get name of datatype:
        //	sDataType := fbJsonDataType.GetDatatypeNameByAddress(			nData        := SIZEOF(CNCSystem.Channel[nChanIdx].ToolData.stOldTool), 
		//  pData        := ADR(CNCSystem.Channel[nChanIdx].ToolData.stOldTool));
			
		// Reset the internal buffer of the JSON writer
    	fbJsonWriter.ResetDocument();
		
		// Serialize the structure into the JSON writer
    	fbJsonDataType.AddJsonValueFromSymbol(
			fbWriter 	 := fbJsonWriter, 
			sDatatype    := 'Tc3_CNC.ST_CNC_TOOL_DATA_EXT', 
			nData        := SIZEOF(CNCSystem.Channel[nChanIdx].ToolData.stOldTool), 
			pData        := ADR(CNCSystem.Channel[nChanIdx].ToolData.stOldTool)
		);
		
		    // Extract the JSON content as a string
    	fbJsonWriter.CopyDocument(
       		pDoc := CNCSystem.Channel[nChanIdx].ToolDataJson.stOldToolJson, 
        	nDoc := SIZEOF(CNCSystem.Channel[nChanIdx].ToolDataJson.stOldToolJson)
   		);
		
		
		IF CNCSystem.Channel[nChanIdx].ToolDataJson.PostToolToJsonAction <> 0 THEN
			nStateOt := nStateOt + 10;   // call ITF action to allow changing the json data
		ELSE
			nStateOt := nStateOt + 20;  // go on directly without calling ITF Action
		END_IF
		
	20: // call ITF Action
		IF CNCSystem.Channel[nChanIdx].ToolDataJson.PostToolToJsonAction.Commit(CNCSystem.Channel[nChanIdx].ToolDataJson.stOldToolJson) THEN
			CNCSystem.Channel[nChanIdx].ToolDataJson.stOldToolJson := CNCSystem.Channel[nChanIdx].ToolDataJson.PostToolToJsonAction.ToolJson;
			nStateOt := nStateOt + 10;
		END_IF

	30:
	
		CNCSystem.Channel[nChanIdx].ToolDataJson.bOldToolDataExist := TRUE;
		nStateOt := nStateOt + 10;		

	40: 
		IF (CNCSystem.Channel[nChanIdx].ToolDataJson.bOldToolDataExist = FALSE) THEN
			nStateOt  := 0;
			CNCSystem.Channel[nChanIdx].ToolData.bOldToolDataExist := FALSE;
		END_IF
		
		 
	
		
END_CASE
END_ACTION

ACTION d_EditToolExists:

CASE nStateEt OF
	
	10:   // forward request to json DataStructure
		  // convert Data to json datastructure			
		  // Reset the internal buffer of the JSON writer
    	fbJsonWriter.ResetDocument();
		
		// Serialize the structure into the JSON writer
    	fbJsonDataType.AddJsonValueFromSymbol(
			fbWriter 	 := fbJsonWriter, 
			sDatatype    := 'Tc3_CNC.ST_CNC_TOOL_DATA_EXT', 
			nData        := SIZEOF(CNCSystem.Channel[nChanIdx].ToolData.stEditTool), 
			pData        := ADR(CNCSystem.Channel[nChanIdx].ToolData.stEditTool)
		);
		
		// Extract the JSON content as a string
    	fbJsonWriter.CopyDocument(
       		pDoc := CNCSystem.Channel[nChanIdx].ToolDataJson.stEditToolJson, 
        	nDoc := SIZEOF(CNCSystem.Channel[nChanIdx].ToolDataJson.stEditToolJson)
   		);
		
		IF CNCSystem.Channel[nChanIdx].ToolDataJson.PostToolToJsonAction <> 0 THEN
			nStateEt := nStateEt + 10;   // call ITF action to allow changing the json data
		ELSE
			nStateEt := nStateEt + 20;  // go on directly without calling ITF Action
		END_IF
		
	20: // call ITF Action
		IF CNCSystem.Channel[nChanIdx].ToolDataJson.PostToolToJsonAction.Commit(CNCSystem.Channel[nChanIdx].ToolDataJson.stEditToolJson) THEN
			CNCSystem.Channel[nChanIdx].ToolDataJson.stEditToolJson := CNCSystem.Channel[nChanIdx].ToolDataJson.PostToolToJsonAction.ToolJson;
			nStateEt := nStateEt + 10;
		END_IF

	30:	
		CNCSystem.Channel[nChanIdx].ToolDataJson.bEditToolDataExist := TRUE;
		nStateEt := nStateEt + 10;		

	40: 
		IF (CNCSystem.Channel[nChanIdx].ToolDataJson.bEditToolDataExist = FALSE) THEN
			nStateEt  := 0;
			CNCSystem.Channel[nChanIdx].ToolData.bEditToolDataExist := FALSE;
		END_IF				 	
		
END_CASE
END_ACTION

METHOD PRIVATE SetSymbolFromJson : BOOL
VAR_INPUT
	jsonDoc : SJsonValue;
	toolData: POINTER TO ST_CNC_TOOL_DATA_EXT;
END_VAR
VAR
	toolDescObj : SJsonValue;
	toolIdObj : SJsonValue;
	toolLifeObj : SJsonValue;
	arrVal : SJsonValue;
	i : INT;
END_VAR
// Top-level fields
toolData^.descriptionText := fbJsonParser.GetString(fbJsonParser.FindMember(jsonDoc, 'descriptionText'));
toolData^.dist_max := fbJsonParser.GetInt(fbJsonParser.FindMember(jsonDoc, 'dist_max'));
toolData^.laenge := fbJsonParser.GetInt(fbJsonParser.FindMember(jsonDoc, 'laenge'));
toolData^.laenge_delta := fbJsonParser.GetInt(fbJsonParser.FindMember(jsonDoc, 'laenge_delta'));
toolData^.pos := fbJsonParser.GetInt(fbJsonParser.FindMember(jsonDoc, 'pos'));
toolData^.radius := fbJsonParser.GetInt(fbJsonParser.FindMember(jsonDoc, 'radius'));
toolData^.radius_delta := fbJsonParser.GetInt(fbJsonParser.FindMember(jsonDoc, 'radius_delta'));
toolData^.time_max := fbJsonParser.GetInt(fbJsonParser.FindMember(jsonDoc, 'time_max'));
toolData^.toleranceNeg := fbJsonParser.GetInt(fbJsonParser.FindMember(jsonDoc, 'toleranceNeg'));
toolData^.tolerancePos := fbJsonParser.GetInt(fbJsonParser.FindMember(jsonDoc, 'tolerancePos'));

// tool_desc object
toolDescObj := fbJsonParser.FindMember(jsonDoc, 'tool_desc');
IF toolDescObj <> 0 THEN
	
	// tool_id object
	toolIdObj := fbJsonParser.FindMember(toolDescObj, 'tool_id');
	IF toolIdObj <> 0 THEN
		toolData^.tool_desc.tool_id.basic := fbJsonParser.GetInt(fbJsonParser.FindMember(toolIdObj, 'basic'));
		toolData^.tool_desc.tool_id.sister := fbJsonParser.GetInt(fbJsonParser.FindMember(toolIdObj, 'sister'));
		toolData^.tool_desc.tool_id.sister_valid := fbJsonParser.GetBool(fbJsonParser.FindMember(toolIdObj, 'sister_valid'));
		toolData^.tool_desc.tool_id.variant := fbJsonParser.GetInt(fbJsonParser.FindMember(toolIdObj, 'variant'));
		toolData^.tool_desc.tool_id.variant_valid := fbJsonParser.GetBool(fbJsonParser.FindMember(toolIdObj, 'variant_valid'));
	END_IF


	toolData^.tool_desc.a_max := fbJsonParser.GetDouble(fbJsonParser.FindMember(toolDescObj, 'a_max'));
	toolData^.tool_desc.additional_settings := UDINT_TO_USINT(fbJsonParser.GetUint(fbJsonParser.FindMember(toolDescObj, 'additional_settings')));
	toolData^.tool_desc.disc_min_radius := fbJsonParser.GetDouble(fbJsonParser.FindMember(toolDescObj, 'disc_min_radius'));
	toolData^.tool_desc.disc_min_width := fbJsonParser.GetDouble(fbJsonParser.FindMember(toolDescObj, 'disc_min_width'));
	toolData^.tool_desc.disc_tilt_angle := fbJsonParser.GetDouble(fbJsonParser.FindMember(toolDescObj, 'disc_tilt_angle'));
	toolData^.tool_desc.ext_discret_limit := fbJsonParser.GetDouble(fbJsonParser.FindMember(toolDescObj, 'ext_discret_limit'));
	toolData^.tool_desc.gear_inv_direction := fbJsonParser.GetBool(fbJsonParser.FindMember(toolDescObj, 'gear_inv_direction'));
	toolData^.tool_desc.gear_inv_direction_no_stop := fbJsonParser.GetBool(fbJsonParser.FindMember(toolDescObj, 'gear_inv_direction_no_stop'));
	toolData^.tool_desc.gear_ratio_denom := fbJsonParser.GetInt(fbJsonParser.FindMember(toolDescObj, 'gear_ratio_denom'));
	toolData^.tool_desc.gear_ratio_num := fbJsonParser.GetInt(fbJsonParser.FindMember(toolDescObj, 'gear_ratio_num'));
	toolData^.tool_desc.kin_id := UDINT_TO_UINT(fbJsonParser.GetUint(fbJsonParser.FindMember(toolDescObj, 'kin_id')));
	toolData^.tool_desc.laenge := fbJsonParser.GetInt(fbJsonParser.FindMember(toolDescObj, 'laenge'));
	toolData^.tool_desc.log_ax_nr_spdl := UDINT_TO_UINT(fbJsonParser.GetUInt(fbJsonParser.FindMember(toolDescObj, 'log_ax_nr_spdl')));
	toolData^.tool_desc.mass_einheit := UDINT_TO_UINT(fbJsonParser.GetUInt(fbJsonParser.FindMember(toolDescObj, 'mass_einheit')));
	toolData^.tool_desc.radius := fbJsonParser.GetInt(fbJsonParser.FindMember(toolDescObj, 'radius'));
	toolData^.tool_desc.radius_path2 := fbJsonParser.GetInt(fbJsonParser.FindMember(toolDescObj, 'radius_path2'));
	toolData^.tool_desc.srk_lage := UDINT_TO_UINT(fbJsonParser.GetUInt(fbJsonParser.FindMember(toolDescObj, 'srk_lage')));
	toolData^.tool_desc.tool_fixed := fbJsonParser.GetBool(fbJsonParser.FindMember(toolDescObj, 'tool_fixed'));
	toolData^.tool_desc.tool_sub_type := UDINT_TO_UINT(fbJsonParser.GetUInt(fbJsonParser.FindMember(toolDescObj, 'tool_sub_type')));
	toolData^.tool_desc.typ := UDINT_TO_UINT(fbJsonParser.GetUInt(fbJsonParser.FindMember(toolDescObj, 'typ')));
	toolData^.tool_desc.valid := fbJsonParser.GetBool(fbJsonParser.FindMember(toolDescObj, 'valid'));
	toolData^.tool_desc.vb_max := fbJsonParser.GetDouble(fbJsonParser.FindMember(toolDescObj, 'vb_max'));
	toolData^.tool_desc.vb_min := fbJsonParser.GetDouble(fbJsonParser.FindMember(toolDescObj, 'vb_min'));
	toolData^.tool_desc.wear_const := fbJsonParser.GetDouble(fbJsonParser.FindMember(toolDescObj, 'wear_const'));

	// add_info array [2]
	arrVal := fbJsonParser.FindMember(toolDescObj, 'add_info');
	IF arrVal <> 0 THEN
		FOR i := 0 TO 1 DO
			toolData^.tool_desc.add_info[i] := DINT_TO_DWORD(fbJsonParser.GetInt(fbJsonParser.GetArrayValueByIdx(arrVal, DINT_TO_UDINT(i))));
		END_FOR
	END_IF

	// ax_versatz array [32]
	arrVal := fbJsonParser.FindMember(toolDescObj, 'ax_versatz');
	IF arrVal <> 0 THEN
		FOR i := 0 TO 31 DO
			toolData^.tool_desc.ax_versatz[i] := fbJsonParser.GetInt(fbJsonParser.GetArrayValueByIdx(arrVal, DINT_TO_UDINT(i)));
		END_FOR
	END_IF

	// kopf_versatz array [70]
	arrVal := fbJsonParser.FindMember(toolDescObj, 'kopf_versatz');
	IF arrVal <> 0 THEN
		FOR i := 0 TO 69 DO
			toolData^.tool_desc.kopf_versatz[i] := fbJsonParser.GetInt(fbJsonParser.GetArrayValueByIdx(arrVal, DINT_TO_UDINT(i)));
		END_FOR
	END_IF

	// orientation_vector array [3]
	arrVal := fbJsonParser.FindMember(toolDescObj, 'orientation_vector');
	IF arrVal <> 0 THEN
		FOR i := 0 TO 2 DO
			toolData^.tool_desc.orientation_vector[i] := fbJsonParser.GetDouble(fbJsonParser.GetArrayValueByIdx(arrVal, DINT_TO_UDINT(i)));
		END_FOR
	END_IF

	// param array [60]
	arrVal := fbJsonParser.FindMember(toolDescObj, 'param');
	IF arrVal <> 0 THEN
		FOR i := 0 TO 59 DO
			toolData^.tool_desc.param[i] := fbJsonParser.GetDouble(fbJsonParser.GetArrayValueByIdx(arrVal, DINT_TO_UDINT(i)));
		END_FOR
	END_IF


END_IF

// tool_life object
toolLifeObj := fbJsonParser.FindMember(jsonDoc, 'tool_life');
IF toolLifeObj <> 0 THEN
	toolData^.tool_life.dist_used := fbJsonParser.GetDouble(fbJsonParser.FindMember(toolLifeObj, 'dist_used'));
	toolData^.tool_life.time_used := fbJsonParser.GetDouble(fbJsonParser.FindMember(toolLifeObj, 'time_used'));
END_IF

SetSymbolFromJson := TRUE;
END_METHOD

END_FUNCTION_BLOCK

// CNC/8 Mis/HLI3_SetPLCAlive
FUNCTION HLI3_SetPLCAlive : BOOL
VAR_INPUT
	nChanIdx: INT;		
END_VAR

VAR
	nWatchdogCycles 	: UDINT :=2;	 	
END_VAR

(*
Display PLC is just alive (Trigger Watchdog to MC)
If PLC is stopped here, alive sign is missing.
-> CNC raises error message
-> CNC stoppes movement with internal FEEDHOLD
-> system has to be restarted (after removal of error)
*)

HLI3_SetPLCAlive := FALSE;
IF NOT HLI3_CheckChannelValid(nChannel := nChanIdx) THEN
	RETURN;
END_IF

nWatchdogCycles := 8;

gpCh[nChanIdx]^.head.mc_watchdog.cycle_time_w := CNCSystem.nPLCCycleTime * nWatchdogCycles;   // Watchdog time : PLC Cycle Time * nWatchdogCycles
gpCh[nChanIdx]^.head.mc_watchdog.enable_w := TRUE;
gpCh[nChanIdx]^.head.mc_watchdog.alive_rw := TRUE;

HLI3_SetPLCAlive := TRUE;

END_FUNCTION

// CNC/3 Control/HLI3_ChannelSetEmergencyStop
FUNCTION HLI3_ChannelSetEmergencyStop : BOOL
VAR_INPUT
	/// Number of channel 
	nChanIdx: INT;
	bEStop: BOOL;
END_VAR

(****************************************************************************************)
(* POU:			HLI_ChannelSetEmergenyStop												*)
(* Type:		Function block															*)
(* Customer:	Common																	*)
(* Date:		09/03/12																*)
(* Last:		20/11/12																*)
(* ------------------------------------------------------------------------------------ *)
(* Revision:	1.0																		*)
(* Author:		HR,MiB																	*)
(* Description: (Re-)Sets the channel specific emergency stop unit.						*)
(****************************************************************************************)

HLI3_ChannelSetEmergencyStop := FALSE;
IF NOT HLI3_CheckChannelValid(nChannel := nChanIdx) THEN
	RETURN;
END_IF

(* if the stop button from the HMI is selected the request is set *)
gpCh[nChanIdx]^.bahn_mc_control.emergency_stop.command_w := bEStop;

HLI3_ChannelSetEmergencyStop		:= TRUE;

END_FUNCTION

// CNC/3 Control/HLI3_SetChannelOverride
FUNCTION HLI3_SetChannelOverride : BOOL
VAR_INPUT
	/// Number of channel 
	nChanIdx: INT;
	nOverride: UINT;
END_VAR

(* ========================================================= *)
(*    FUN: HLI_SetChannelOverride                            *)
(* --------------------------------------------------------- *)
(*   Desc: Set the channel Override                          *)
(* Author: MK, MiB                                           *)
(*   Date: 20.11.2012                                        *)
(*   Rev.: 1.2  2017.10.25                                   *)
(* ========================================================= *)

IF NOT HLI3_CheckChannelValid(nChannel := nChanIdx) THEN
	HLI3_SetChannelOverride := FALSE;
	RETURN;
END_IF

(* Limit the override *)
IF nOverride > 2000 THEN nOverride := 2000; END_IF  // MiB 2017.10.25 valid maximum in cnc core is 2000
IF nOverride < 0 THEN nOverride := 0; END_IF

gpCh[nChanIdx]^.bahn_mc_control.override_feedrate.command_w := nOverride;

HLI3_SetChannelOverride := TRUE;

END_FUNCTION

// CNC/3 Control/HLI3_SetChannelRapidOverride
FUNCTION HLI3_SetChannelRapidOverride : BOOL
VAR_INPUT
	/// Number of channel 
	nChanIdx: INT;
	nOverride: UINT;
END_VAR

(* ========================================================= *)
(*    FUN: HLI_SetChannelRapidOverride                       *)
(* --------------------------------------------------------- *)
(*   Desc: Set the channel Override for rapid movements      *)
(*   Author: TV , MiB                                        *)
(*   Date: 07.02.2017                                        *)
(*   Rev.: 1.1                                               *)
(* ========================================================= *)

IF NOT HLI3_CheckChannelValid(nChannel := nChanIdx) THEN
	HLI3_SetChannelRapidOverride := FALSE;
	RETURN;
END_IF

(* Limit the override *)
IF nOverride > 1000	THEN nOverride := 1000; END_IF  // MiB 2017.10.25 maximum is 1000 (ref HLI manual)
IF nOverride < 0 THEN nOverride := 0; END_IF

gpCh[nChanIdx]^.bahn_mc_control.override_rapid_move.enable_w := TRUE;
gpCh[nChanIdx]^.bahn_mc_control.override_rapid_move.command_w := nOverride;

HLI3_SetChannelRapidOverride := TRUE;

END_FUNCTION

// CNC/3 Control/HLI3_ChannelSetBackwardMotion
FUNCTION HLI3_ChannelSetBackwardMotion : BOOL
VAR_INPUT
	/// Number of channel 
	nChanIdx: INT;
	bBackwardMotion: BOOL;
END_VAR

(* ========================================================= *)
(*    FUN: HLI_ChannelSetBackwardMotion                      *)
(* --------------------------------------------------------- *)
(*   Desc:                                                   *)
(* Author: MK, MiB                                           *)
(*   Date: 20.11.2012                                        *)
(*   Rev.: 1.1                                               *)
(* ========================================================= *)

HLI3_ChannelSetBackwardMotion := FALSE;
IF NOT HLI3_CheckChannelValid(nChannel := nChanIdx) THEN
	RETURN;
END_IF

gpCh[nChanIdx]^.bahn_mc_control.backward_motion.command_w := bBackwardMotion;

HLI3_ChannelSetBackwardMotion := TRUE;

END_FUNCTION

// CNC/3 Control/HLI3_ChannelSetProgramBlockIgnore
FUNCTION HLI3_ChannelSetProgramBlockIgnore : BOOL
VAR_INPUT
	/// Number of channel 
	nChanIdx: INT;
	bPrgBlockIgnore: BOOL;
END_VAR

(* ========================================================= *)
(*    FUN: HLI_SetProgramBlockIgnore                         *)
(* --------------------------------------------------------- *)
(*   Desc:                                                   *)
(* Author: MK, MiB , TV                                      *)
(*   Date: 20.12.2012                                        *)
(*   Last: 19.11.2013                                        *)
(*   Rev.: 1.0                                               *)
(* ========================================================= *)

HLI3_ChannelSetProgramBlockIgnore := FALSE;
IF NOT HLI3_CheckChannelValid(nChannel := nChanIdx) THEN
	RETURN;
END_IF

(* program block ignore *)
IF bPrgBlockIgnore THEN
	gpCh[nChanIdx]^.decoder_mc_control.program_block_ignore.command_w := 1;
ELSE
	gpCh[nChanIdx]^.decoder_mc_control.program_block_ignore.command_w := 0;
END_IF

HLI3_ChannelSetProgramBlockIgnore := TRUE;

END_FUNCTION

// CNC/3 Control/HLI3_ChannelSetFeedHold
FUNCTION HLI3_ChannelSetFeedHold : BOOL
VAR_INPUT
	/// Number of channel 
	nChanIdx: INT;
	bFeedHold: BOOL;
END_VAR

(* ========================================================= *)
(*    FUN: HLI_ChannelSetFeedHold                            *)
(* --------------------------------------------------------- *)
(*   Desc:                                                   *)
(* Author: MK , MiB                                          *)
(*   Date: 20.11.2012                                        *)
(*   Rev.: 1.1                                               *)
(* ========================================================= *)

HLI3_ChannelSetFeedHold := FALSE;
IF NOT HLI3_CheckChannelValid(nChannel := nChanIdx) THEN
	RETURN;
END_IF

(* if the stop button from the HMI is selected the request is set *)
gpCh[nChanIdx]^.bahn_mc_control.feedhold.command_w := bFeedHold OR gpCh[nChanIdx]^.bahn_mc_control.feedhold.request_r;
HLI3_ChannelSetFeedHold := TRUE;

END_FUNCTION

// CNC/3 Control/HLI3_ChannelSetSingleBlock
FUNCTION HLI3_ChannelSetSingleBlock : BOOL
VAR_INPUT
	/// Number of channel 
	nChanIdx: INT;
	bSingleBlock: BOOL;
END_VAR

(* ========================================================= *)
(*    FUN: HLI3_ChannelSetSingleBlock                        *)
(* --------------------------------------------------------- *)
(*   Desc:                                                   *)
(* Author: MK ,MiB                                           *)
(*   Date: 20.11.2012                                        *)
(*   Rev.: 1.1                                               *)
(* ========================================================= *)

HLI3_ChannelSetSingleBlock := FALSE;
IF NOT HLI3_CheckChannelValid(nChannel := nChanIdx) THEN
	RETURN;
END_IF
gpCh[nChanIdx]^.bahn_mc_control.single_block.command_w   := bSingleBlock;

HLI3_ChannelSetSingleBlock := TRUE;

END_FUNCTION

// CNC/3 Control/HLI3_ChannelSetReducedFeed
FUNCTION HLI3_ChannelSetReducedFeed : BOOL
VAR_INPUT
	/// Number of channel 
	nChanIdx: INT;
	bReducedFeed: BOOL;
END_VAR

(* ========================================================= *)
(*    FUN: HLI_ChannelSetReducedFeed                         *)
(* --------------------------------------------------------- *)
(*   Desc:                                                   *)
(* Author: MK,MiB                                            *)
(*   Date: 20.11.2012                                        *)
(*   Rev.: 1.1                                               *)
(* ========================================================= *)


HLI3_ChannelSetReducedFeed := FALSE;
IF NOT HLI3_CheckChannelValid(nChannel := nChanIdx) THEN
	RETURN;
END_IF
gpCh[nChanIdx]^.bahn_mc_control.reduced_speed.command_w := bReducedFeed;
HLI3_ChannelSetReducedFeed := TRUE;

END_FUNCTION

// CNC/3 Control/HLI3_GetChannelStatusInfo
FUNCTION HLI3_GetChannelStatusInfo : BOOL
VAR_INPUT
	/// Number of channel 
	nChanIdx: INT;
END_VAR
VAR
	pChannel: POINTER TO ST_CNCChannel;
END_VAR

(* ========================================================= *)
(*    FUN: HLI_GetStatusInfo                                 *)
(* --------------------------------------------------------- *)
(*   Desc: Status Info from the HLI Interface                *)
(* Author: MK,Mib                                            *)
(*   Date: 18.07.2002                                        *)
(*   Rev.: 1.0                                               *)
(* ========================================================= *)

IF NOT HLI3_CheckChannelValid(nChannel := nChanIdx) THEN
	RETURN;
END_IF


pChannel := ADR(CNCSystem.Channel[nChanIdx]);
pChannel^.ActMode := HLI3_GetChannelMode(nChanIdx:=nChanIdx);
pChannel^.ActState := HLI3_GetChannelState(nChanIdx:=nChanIdx);

pChannel^.Mode.Standby := FALSE;
pChannel^.Mode.Auto := FALSE;
pChannel^.Mode.Homing := FALSE;
pChannel^.Mode.MDI := FALSE;
pChannel^.Mode.Manual := FALSE;

(* Translate mode *)
CASE pChannel^.ActMode OF
	HLI_IMCM_MODE:					pChannel^.ActModeString := 'Mode';
	HLI_IMCM_STANDBY_MODE:			pChannel^.ActModeString := 'StandbyMode'; pChannel^.Mode.Standby:=TRUE;
	HLI_IMCM_AUTOMATIC_MODE:		pChannel^.ActModeString := 'AutomaticMode'; pChannel^.Mode.Auto:=TRUE;
	HLI_IMCM_MDI_MODE:				pChannel^.ActModeString := 'MDIMode'; pChannel^.Mode.MDI:=TRUE;
	HLI_IMCM_MANUAL_MODE:			pChannel^.ActModeString := 'ManualMode'; pChannel^.Mode.Manual:=TRUE;;
	HLI_IMCM_REFERENCE_MODE:		pChannel^.ActModeString := 'ReferenceMode'; pChannel^.Mode.Homing:=TRUE;
ELSE
	pChannel^.ActModeString := '---';
END_CASE;

pChannel^.State.Selected:=FALSE;
pChannel^.State.Ready:=FALSE;
pChannel^.State.Active:=FALSE;
pChannel^.State.Hold:=FALSE;
pChannel^.State.Error:=FALSE;

(* Translate state *)
CASE pChannel^.ActState OF
	HLI_IMCM_PROCESS_DESELECTED:	pChannel^.ActStateString := 'Deselected';
	HLI_IMCM_PROCESS_SELECTED:		pChannel^.ActStateString := 'Selected'; pChannel^.State.Selected:=TRUE;
	HLI_IMCM_PROCESS_READY:			pChannel^.ActStateString := 'Ready'; pChannel^.State.Ready:=TRUE;
	HLI_IMCM_PROCESS_ACTIVE:		pChannel^.ActStateString := 'Active'; pChannel^.State.Active:=TRUE;
	HLI_IMCM_PROCESS_HOLD:			pChannel^.ActStateString := 'Hold'; pChannel^.State.Hold:=TRUE;
	HLI_IMCM_PROCESS_ERROR:			pChannel^.ActStateString := 'Error'; pChannel^.State.Error:=TRUE;
	HLI_IMCM_PROCESS_SELECTING:		pChannel^.ActStateString := 'Selecting';
	HLI_IMCM_PROCESS_DESELECTING:	pChannel^.ActStateString := 'Deselecting';
	HLI_IMCM_PROCESS_PREPARING:		pChannel^.ActStateString := 'Preparing';
	HLI_IMCM_PROCESS_CLEARING:		pChannel^.ActStateString := 'Clearing';
	HLI_IMCM_PROCESS_STARTING:		pChannel^.ActStateString := 'Starting';
	HLI_IMCM_PROCESS_ABORTING:		pChannel^.ActStateString := 'Aborting';
	HLI_IMCM_PROCESS_STOPPING:		pChannel^.ActStateString := 'Stopping';
	HLI_IMCM_PROCESS_RESUMING:		pChannel^.ActStateString := 'Resuming';
	HLI_IMCM_PROCESS_RESETTING:		pChannel^.ActStateString := 'Resetting';
	HLI_IMCM_PROCESS_FINISHING:		pChannel^.ActStateString := 'Finishing';
ELSE
	pChannel^.ActStateString := '---';
END_CASE;

END_FUNCTION

// CNC/3 Control/HLI3_GetChannelMode
FUNCTION HLI3_GetChannelMode : UDINT
VAR_INPUT
	/// Number of channel 
	nChanIdx: INT;
END_VAR

(* ========================================================= *)
(*    FUN: HLI_GetChannelMode                                *)
(* --------------------------------------------------------- *)
(*   Desc:                                                   *)
(* Author: MK                                                *)
(*   Date: 18.07.2002                                        *)
(*   Rev.: 1.0                                               *)
(* ========================================================= *)
HLI3_GetChannelMode := 0;
IF NOT HLI3_CheckChannelValid(nChannel := nChanIdx) THEN
	RETURN;
END_IF

(* if the stop button from the HMI is selected the request is set *)
HLI3_GetChannelMode := gpCh[nChanIdx]^.channel_mc_control.mode_and_state.state_r.mode;

END_FUNCTION

// CNC/3 Control/HLI3_GetChannelState
FUNCTION HLI3_GetChannelState : UDINT
VAR_INPUT
	/// Number of channel 
	nChanIdx: INT;
END_VAR

(* ========================================================= *)
(*    FUN: HLI3_GetChannelState                              *)
(* --------------------------------------------------------- *)
(*   Desc:                                                   *)
(* Author: MK                                                *)
(*   Date: 18.07.2002                                        *)
(*   Rev.: 1.0                                               *)
(* ========================================================= *)

HLI3_GetChannelState := 0;
IF NOT HLI3_CheckChannelValid(nChannel := nChanIdx) THEN
	RETURN;
END_IF

(* if the stop button from the HMI is selected the request is set *)
HLI3_GetChannelState := gpCh[nChanIdx]^.channel_mc_control.mode_and_state.state_r.state;

END_FUNCTION

// CNC/3 Control/HLI3_GetChannelError
FUNCTION HLI3_GetChannelError : BOOL
VAR_INPUT
	/// Number of channel 
	nChanIdx: INT;
END_VAR
VAR
	pChannel: POINTER TO ST_CNCChannel;
END_VAR

(* ========================================================= *)
(*    FUN: HLI_GetChannelError                               *)
(* --------------------------------------------------------- *)
(*   Desc: Gets the channel error                            *)
(* Return: The error flag of the channel                     *)
(* Author: MK , MiB, TV                                      *)
(*   Date: 25.10.2023                                        *)
(*   Rev.: 1.4                                               *)
(* ========================================================= *)

IF NOT HLI3_CheckChannelValid(nChannel := nChanIdx) THEN
	RETURN;
END_IF

pChannel := ADR(CNCSystem.Channel[nChanIdx]);

(* Visualisation of Mode and State *)
pChannel^.ActMode  := HLI3_GetChannelMode(nChanIdx:=nChanIdx);
pChannel^.ActState := HLI3_GetChannelState(nChanIdx:=nChanIdx);

(* Error messages id *)
IF pChannel^.ActState = HLI_IMCM_PROCESS_ERROR THEN
	pChannel^.Error := TRUE;	
	HLI3_GetChannelError := TRUE;
ELSE
	pChannel^.Error := FALSE;	
	HLI3_GetChannelError := FALSE;
END_IF

END_FUNCTION

// CNC/4 MHT-Function/HLI3_QuitChannelMHTFunction
FUNCTION_BLOCK HLI3_QuitChannelMHTFunction
VAR_INPUT
	/// Number of channel 
	nChanIdx: INT;
	bM30Acknowledgement : BOOL;
	bDisableAutoAcknowledgeM : BOOL;
END_VAR
VAR_OUTPUT
	bOK: BOOL;
END_VAR
VAR
	ChannelMFunction: HLI3_DoChannelMFunction;
	ChannelMFunctionLateSync : HLI3_DoChannelMFunction;
	ChannelTFunction: HLI3_DoChannelTFunction;
	ChannelHFunction: HLI3_DoChannelHFunction;
	/// local pointer to Data of actual Channel 
	pChannelData: POINTER TO HIGH_LEVEL_INTERFACE_CH;
	/// local pointer to actual techno unit 
	pActTechnoUnit: POINTER TO TECHNO_UNIT_CH;
	/// Index of axis specific technology function at HLI 
	nTechFctMaxIdx: UINT;
	nTechFctAnzahl : UINT; 
	/// loop variable 
	idx: UINT;
	/// number of M-function 
	nFuncNr: UDINT;
	nArgument: DINT;
	/// basis id of a tool 
	nToolBasicId: UDINT;
	pMHProcess: POINTER TO HLI_M_H_PROZESS;
	pSProcess: POINTER TO HLI_S_PROZESS;
	pTProcess: POINTER TO HLI_T_PROZESS;
	stAttributeData: St_TechnoAttributeData;	
END_VAR

(* ========================================================= *)
(*     FB: HLI3_QuitChannelMHTFunction                        *)
(* --------------------------------------------------------- *)
(*   Desc:                                                   *)
(* Author: MK                                                *)
(*   Rev.: 1.1                                               *)
(*   Date: 18.07.2002                                        *)
(*       : 08.04.2005                                        *)
(*          24.11.2010 MiB Erweiterung um H Funktionen 		 *)
(* ========================================================= *)
(* Rev.:	1.2												 *)
(* Date:	02.10.2010                                    	 *)
(* Author:	HR												 *)
(* Author:	Added support for additional m function number	 *)
(* ========================================================= *)
(* Rev.:	1.3												 *)
(* Date:	26.01.2011                                    	 *)
(* Author:	HR												 *)
(* Author:	Added support for additional h function number	 *)
(* ========================================================= *)
(* Rev.:	1.4												 *)
(* Date:	20.11.2012                                    	 *)
(* Author:	MiB												 *)
(* Author:	TC3												 *)
(* ========================================================= *)
(* Rev.:	1.4.1									         *)
(* Date:	15.07.2013                                    	 *)
(* Author:	TV												 *)
(* ========================================================= *)
(* Rev.:	1.4.2									         *)
(* Date:	22.09.2016                                    	 *)
(* Author:	TV												 *)
(* ========================================================= *)
(* ========================================================= *)
(* Rev.:	1.4.3									         *)
(* Date:	01.12.2017                                    	 *)
(* Author:	TV												 *)
(*													 	 	 *)
(* ========================================================= *)

IF NOT HLI3_CheckChannelValid(nChannel := nChanIdx) THEN
	bOK := FALSE;
	RETURN; (* A b b r u c h *)
END_IF


(* get pointer to channel data *)
pChannelData := gpCh[nChanIdx];

pActTechnoUnit := ADR(pChannelData^.techno_unit_std_sync[0]);

(* test if there are open synchronisations  *)
IF pChannelData^.used_units_std_sync_r > 0 THEN

	nTechFctAnzahl := pChannelData^.used_units_std_sync_r;
	
	IF nTechFctAnzahl  > 0 THEN

        nTechFctMaxIdx := nTechFctAnzahl  - 1;  

		FOR idx := 0 TO nTechFctMaxIdx DO
			(* get pointer to actual techno unit *)
			pActTechnoUnit := ADR(pChannelData^.techno_unit_std_sync[idx]);
		
		
			(* test if this M-function has to be acknowledged *)
			IF pActTechnoUnit^.please_rw = TRUE AND				(* request from CNC *)
			   pActTechnoUnit^.done_w = FALSE AND				(* not acknowledged *)
			   pActTechnoUnit^.fkt_ctrl_r = HLI_INTF_M_FKT		(* M-function *)
			THEN
				(* Read number of M-function *)
				pMHProcess := ADR(pActTechnoUnit^.attribut_r.data[0]);
				nFuncNr    := pMHProcess^.nr;
				nArgument	:= pMHProcess^.add_nr_r;
				
				
				stAttributeData.nFunctionNumber_r := pMHProcess^.nr;
				stAttributeData.nTime_r		:= pMHProcess^.zeit;
				stAttributeData.nArgument_r 		:= pMHProcess^.add_nr_r;
				stAttributeData.nBlockNumber_r 	:= pMHProcess^.satz_nr;
				stAttributeData.nPrgLineNumber_r	:= pMHProcess^.prg_zeilen_nr;
				
		
				ChannelMFunction(nChanIdx:=nChanIdx, stTechnoAttributeData := stAttributeData, bM30Acknowledgement := bM30Acknowledgement, bDisableAutoAcknowledgeM := bDisableAutoAcknowledgeM);
				IF ChannelMFunction.bBusy = FALSE THEN
					(* acknowledge this M-function *)
					pActTechnoUnit^.please_rw := FALSE;
					pActTechnoUnit^.done_w := TRUE;				
				END_IF
		
				bOK := TRUE;
			END_IF
	
	
			(* test if this H-function has to be acknowledged *)
			IF pActTechnoUnit^.please_rw = TRUE AND						(* request from CNC *)
			   pActTechnoUnit^.done_w = FALSE AND						(* not acknowledged *)
			   pActTechnoUnit^.fkt_ctrl_r = HLI_INTF_H_FKT		(* H-function *)
			THEN
				(* Read number of H-function *)
				pMHProcess := ADR(pActTechnoUnit^.attribut_r.data[0]);
				stAttributeData.nFunctionNumber_r := pMHProcess^.nr;
				stAttributeData.nTime_r		:= pMHProcess^.zeit;
				stAttributeData.nArgument_r 		:= pMHProcess^.add_nr_r;
				stAttributeData.nBlockNumber_r 	:= pMHProcess^.satz_nr;
				stAttributeData.nPrgLineNumber_r	:= pMHProcess^.prg_zeilen_nr;
		
				ChannelHFunction(nChanIdx:=nChanIdx, stTechnoAttributeData:= stAttributeData);
	
				(* acknowledge this H-function *)
				IF ChannelHFunction.bBusy = FALSE THEN
						(* acknowledge this H-function *)
					pActTechnoUnit^.please_rw := FALSE;
					pActTechnoUnit^.done_w := TRUE;			
				END_IF
				bOK := TRUE;
			END_IF
		
			(* test if this T-function has to be acknowledged *)
			IF pActTechnoUnit^.please_rw = TRUE AND				(* request from CNC *)
			   pActTechnoUnit^.done_w = FALSE AND				(* not acknowledged *)
			   pActTechnoUnit^.fkt_ctrl_r = HLI_INTF_TOOL		(* T-function *)
			THEN
				(* Read number of T-function *)
				pTProcess    := ADR(pActTechnoUnit^.attribut_r.data[0]);
				nToolBasicId := DINT_TO_UDINT(pTProcess^.id.basic);
		
				ChannelTFunction(nChanIdx:=nChanIdx, nFuncNr:=nToolBasicId);
		
				(* acknowledge this T-function *)
				pActTechnoUnit^.please_rw := FALSE;
				pActTechnoUnit^.done_w := TRUE;				
				bOK := TRUE;
			END_IF
		
		END_FOR
	
	END_IF

END_IF


(*
	HLI_INTF_H_FKT                 :    INT:=2;
	HLI_INTF_SPINDEL              :    INT:=3;
	HLI_INTF_TOOL                 :    INT:=4;
	GCW_250_HLIIntfAxBlock              :    INT:=5;
	GCW_250_HLIIntfVEVariable           :    INT:=6;
	GCW_250_HLIIntfVEVariable_1         :    INT:=7;
	GCW_250_HLIIntfVEVariable_2         :    INT:=8;
	GCW_250_HLIIntfUnknown              :    INT:=9;
*)

(*******************************************************************************************************************)

FOR idx := 0 TO INT_TO_UINT(HLI_TU_CH_LATE_SYNC_MAXIDX) DO
	IF pChannelData^.techno_unit_late_sync[idx].please_rw = TRUE
	AND pChannelData^.techno_unit_late_sync[idx].done_w = FALSE THEN

		(* get pointer to actual techno unit *)
		pActTechnoUnit := ADR(pChannelData^.techno_unit_late_sync[idx]);

		IF pActTechnoUnit^.please_rw = TRUE AND				(* request from CNC *)
			pActTechnoUnit^.done_w = FALSE AND				(* not acknowledged *)
			pActTechnoUnit^.fkt_ctrl_r = HLI_INTF_M_FKT		(* M-function *)
		THEN
			pMHProcess := ADR(pActTechnoUnit^.attribut_r.data[0]);
			nFuncNr    := pMHProcess^.nr;
			
			stAttributeData.nFunctionNumber_r := pMHProcess^.nr;
			stAttributeData.nTime_r		:= pMHProcess^.zeit;
			stAttributeData.nArgument_r 		:= pMHProcess^.add_nr_r;
			stAttributeData.nBlockNumber_r 	:= pMHProcess^.satz_nr;
			stAttributeData.nPrgLineNumber_r	:= pMHProcess^.prg_zeilen_nr;

			ChannelMFunctionLateSync(nChanIdx:=nChanIdx, stTechnoAttributeData:=stAttributeData,bM30Acknowledgement := bM30Acknowledgement, bDisableAutoAcknowledgeM := bDisableAutoAcknowledgeM);
			IF ChannelMFunctionLateSync.bBusy = FALSE THEN
				(* acknowledge this M-function *)
				pActTechnoUnit^.please_rw := FALSE;
				pActTechnoUnit^.done_w := TRUE;
				
				(* ADSLOGDINT( msgCtrlMask := ADSLOG_MSGTYPE_MSGBOX OR
											ADSLOG_MSGTYPE_LOG,
							msgFmtStr := 'Channel acknowledge of M-function: %d',
							dintArg := pMHProcess^.nr);
				*)
			END_IF
		bOK := TRUE;

	(*	ELSIF   pActTechnoUnit^.fkt_ctrl_r = HLI_INTF_SPINDEL THEN (* spindle-function *)

 			(* Example: read number of S-function *)
			pSProzess := ADR(pActTechnoUnit^.attribut_r.data[0]);
			ADSLOGDINT( msgCtrlMask := ADSLOG_MSGTYPE_MSGBOX OR
										ADSLOG_MSGTYPE_LOG,
						msgFmtStr := 'Late synch : %d',
						dintArg := pSProzess^.move_cmd);

		ELSIF   pActTechnoUnit^.fkt_ctrl_r = HLI_INTF_TOOL THEN

			pHLI_T_PROZESS := ADR(pActTechnoUnit^.attribut_r.data[0]);
			ADSLOGDINT( msgCtrlMask := ADSLOG_MSGTYPE_MSGBOX OR
										ADSLOG_MSGTYPE_LOG,
						msgFmtStr := 'Late tool process: %d',
						dintArg := pTProcess^.id.basic);*)
		(*ELSE
				ADSLOGDINT( msgCtrlMask := ADSLOG_MSGTYPE_MSGBOX OR
											ADSLOG_MSGTYPE_LOG,
							msgFmtStr := 'Channel acknowledge unknown type: %d',
							dintArg := pActTechnoUnit^.fkt_ctrl_r);*)
		END_IF

	END_IF
END_FOR
(**********************************************************************************************************************)

END_FUNCTION_BLOCK

// CNC/4 MHT-Function/HLI3_DoChannelMFunction
FUNCTION_BLOCK HLI3_DoChannelMFunction
VAR_INPUT
	/// Channel number 
	nChanIdx: INT;
	stTechnoAttributeData: St_TechnoAttributeData;
	bM30Acknowledgement : BOOL;
	bDisableAutoAcknowledgeM : BOOL;  // disable auto acknowledge of M0, M1, M2, M17, M29, M30
END_VAR
VAR_OUTPUT
	bBusy: BOOL;
END_VAR
VAR
	pChannel: POINTER TO ST_CncChannel;
END_VAR

(* ========================================================= *)
(*     FB: HLI_DoChannelMFunction                            *)
(* --------------------------------------------------------- *)
(*   Desc:                                                   *)
(* Author: MK                                                *)
(*   Rev.: 1.1                                               *)
(*   Date: 18.07.2002                                        *)
(*       : 08.04.2005                                        *)
(* ========================================================= *)
(* Rev.:	1.2												 *)
(* Date:	02.10.2010                                   	 *)
(* Author:	HR												 *)
(* Author:	Added support for additional m function number	 *)
(*			via new input variable 'nArg'				 	 *)
(* ========================================================= *)
(* Rev.:	1.3												 *)
(* Date:	23.11.2012                                   	 *)
(* Author:	TV, MiB											 *)
(* Author:	structure St_TechnoAttributeData instead of      *)
(*			simple bool array	 							 *)
(* ========================================================= *)
(* Rev.:	1.4												 *)
(* Date:	22.09.2016                                   	 *)
(* Author:	TV 											 	 *)
(* Dec:		Implementation of Input bM30Acknowledgement      *)
(*				 							                 *)
(* ========================================================= *)

bBusy := TRUE;
IF NOT HLI3_CheckChannelValid(nChannel := nChanIdx) THEN
	RETURN; (* A b b r u c h *)
END_IF


pChannel := ADR(CNCSystem.Channel[nChanIdx]);

(* Synch M-Functions *)
IF stTechnoAttributeData.nFunctionNumber_r >= 0 AND stTechnoAttributeData.nFunctionNumber_r < 1000 THEN
	IF NOT pChannel^.M[stTechnoAttributeData.nFunctionNumber_r].bRes THEN					(* M-Function not set *)		
		pChannel^.M[stTechnoAttributeData.nFunctionNumber_r].nArgument_r		:= stTechnoAttributeData.nArgument_r;
		pChannel^.M[stTechnoAttributeData.nFunctionNumber_r].nBlockNumber_r		:= stTechnoAttributeData.nBlockNumber_r;
		pChannel^.M[stTechnoAttributeData.nFunctionNumber_r].nPrgLineNumber_r	:= stTechnoAttributeData.nPrgLineNumber_r;
		pChannel^.M[stTechnoAttributeData.nFunctionNumber_r].nFunctionNumber_r	:= stTechnoAttributeData.nFunctionNumber_r;
		pChannel^.M[stTechnoAttributeData.nFunctionNumber_r].nTime_r			:= stTechnoAttributeData.nTime_r;		
		pChannel^.M[stTechnoAttributeData.nFunctionNumber_r].bRes 				:= TRUE;	(* set acknowledge *)
		pChannel^.M[stTechnoAttributeData.nFunctionNumber_r].bState_rw			:= TRUE;	(* set M-Function *)
		pChannel^.actM_r := CONCAT('M', UDINT_TO_STRING(stTechnoAttributeData.nFunctionNumber_r));
	ELSE
		IF NOT pChannel^.M[stTechnoAttributeData.nFunctionNumber_r].bState_rw THEN				(* wait for quit *)
			pChannel^.M[stTechnoAttributeData.nFunctionNumber_r].bRes 			:= FALSE;	(* quit the ack *)
			pChannel^.M[stTechnoAttributeData.nFunctionNumber_r].nArgument_r	:= 0;		(* reset the argument *)
			pChannel^.M[stTechnoAttributeData.nFunctionNumber_r].nBlockNumber_r		:= 0;
			pChannel^.M[stTechnoAttributeData.nFunctionNumber_r].nPrgLineNumber_r	:= 0;
			pChannel^.M[stTechnoAttributeData.nFunctionNumber_r].nFunctionNumber_r	:= 0;
			pChannel^.M[stTechnoAttributeData.nFunctionNumber_r].nTime_r			:= 0;				
			pChannel^.actM_r :='';
			bBusy 							:= FALSE;	(* quit *)
		END_IF
	END_IF
END_IF


IF NOT bDisableAutoAcknowledgeM THEN 
	(* Quit M00, M01, M02 , M17, M29, M30 *)
	IF 	stTechnoAttributeData.nFunctionNumber_r = 0 OR 
		stTechnoAttributeData.nFunctionNumber_r = 01 OR 
		stTechnoAttributeData.nFunctionNumber_r = 02 OR 
		stTechnoAttributeData.nFunctionNumber_r = 17  OR 
		stTechnoAttributeData.nFunctionNumber_r = 29  OR 
		(stTechnoAttributeData.nFunctionNumber_r = 30 AND bM30Acknowledgement) THEN
			pChannel^.M[stTechnoAttributeData.nFunctionNumber_r].bState_rw 			:= FALSE;
			pChannel^.M[stTechnoAttributeData.nFunctionNumber_r].nArgument_r	:= 0;
			pChannel^.M[stTechnoAttributeData.nFunctionNumber_r].bRes 			:= FALSE;
			bBusy 							:= FALSE;
	END_IF
END_IF

END_FUNCTION_BLOCK

// CNC/4 MHT-Function/HLI3_DoChannelTFunction
FUNCTION_BLOCK HLI3_DoChannelTFunction
VAR_INPUT
	/// Channel number 
	nChanIdx: INT;
	/// Number of T-function 
	nFuncNr: UDINT;
END_VAR
VAR_OUTPUT
	bBusy: BOOL;
END_VAR
VAR
	bStartTimer: BOOL;
END_VAR

(* ========================================================= *)
(*     FB: HLI_DoChannelTFunction                            *)
(* --------------------------------------------------------- *)
(*   Desc:                                                   *)
(* Author: MK, MiB                                           *)
(*   Rev.: 1.1                                               *)
(*   Date: 18.07.2002                                        *)
(*       : 08.04.2005, 03.03.2016 							 *)
(* ========================================================= *)


bBusy := FALSE;
RETURN;

IF NOT HLI3_CheckChannelValid(nChannel := nChanIdx) THEN
	RETURN; (* A b b r u c h *)
END_IF
bBusy := TRUE;

CASE nChanIdx OF
	0:	(* cnc channel 1 -------------------------------------- *)
		CASE nFuncNr OF
			0:		bBusy := FALSE;
			1:		bBusy := FALSE;
			2:		bBusy := FALSE;
			3:		bBusy := FALSE;
			4:		bBusy := FALSE;
			5:		bBusy := FALSE;
			6:		bBusy := FALSE;
			7:		bBusy := FALSE;
			8:		bBusy := FALSE;

			ELSE
			ADSLOGDINT( msgCtrlMask :=    ADSLOG_MSGTYPE_MSGBOX
			                           OR ADSLOG_MSGTYPE_LOG,
						msgFmtStr   := 'T-Funktion (%d), Channel 1, HLI_DoChannelTFunction() not implemented!',
						dintArg     := UDINT_TO_DINT(nFuncNr));
				(* Quit the M-Function *)
				bBusy := TRUE;
		END_CASE;


	1:	(* cnc channel 2 -------------------------------------- *)
		CASE nFuncNr OF
			0:		bBusy := FALSE;
			1:		bBusy := FALSE;
			2:		bBusy := FALSE;
			3:		bBusy := FALSE;


			ELSE
				ADSLOGDINT( msgCtrlMask :=    ADSLOG_MSGTYPE_MSGBOX
				                           OR ADSLOG_MSGTYPE_LOG,
							msgFmtStr   := 'T-Funktion (%d), Channel 2, HLI_DoChannelTFunction() not implemented!',
							dintArg     := UDINT_TO_DINT(nFuncNr));
				(* Quit the M-Function *)
				bBusy := FALSE;
		END_CASE;

ELSE
	ADSLOGDINT( msgCtrlMask :=    ADSLOG_MSGTYPE_MSGBOX
	                           OR ADSLOG_MSGTYPE_LOG,
				msgFmtStr   := 'Unknown channel number (%d) in HLI_DoChannelTFunction',
				dintArg     := INT_TO_DINT(nChanIdx));
	bBusy := FALSE;
END_CASE;

END_FUNCTION_BLOCK

// CNC/4 MHT-Function/HLI3_DoChannelHFunction
FUNCTION_BLOCK HLI3_DoChannelHFunction
VAR_INPUT
	/// Channel number 
	nChanIdx: INT;
	stTechnoAttributeData: St_TechnoAttributeData;
END_VAR
VAR_OUTPUT
	bBusy: BOOL;
END_VAR
VAR
	pChannel: POINTER TO ST_CncChannel;
END_VAR

(* ========================================================= *)
(*     FB: HLI_DoChannelHFunction                            *)
(* --------------------------------------------------------- *)
(*   Desc:                                                   *)
(* Author: MiB                                               *)
(*   Rev.: 1.0                                               *)
(*   Date: 24.11.2010                                        *)
(*       : 08.04.2005                                        *)
(* ========================================================= *)
(* Rev.:	1.2												 *)
(* Date:	26.01.2011                                   	 *)
(* Author:	HR												 *)
(* Author:	Added support for additional h function number	 *)
(*			via new input variable 'nArg'				 	 *)
(* ========================================================= *)
bBusy := TRUE;

IF NOT HLI3_CheckChannelValid(nChannel := nChanIdx) THEN
	RETURN; (* A b b r u c h *)
END_IF


pChannel := ADR(CNCSystem.Channel[nChanIdx]);

(* Synch M-Functions *)
IF stTechnoAttributeData.nFunctionNumber_r > 0 AND stTechnoAttributeData.nFunctionNumber_r < 1000 THEN
	IF NOT pChannel^.H[stTechnoAttributeData.nFunctionNumber_r].bRes THEN					(* M-Function not set *)
		pChannel^.H[stTechnoAttributeData.nFunctionNumber_r].bState_rw				:= TRUE;	(* set M-Function *)
		pChannel^.H[stTechnoAttributeData.nFunctionNumber_r].nArgument_r		:= stTechnoAttributeData.nArgument_r;
		pChannel^.H[stTechnoAttributeData.nFunctionNumber_r].nBlockNumber_r		:= stTechnoAttributeData.nBlockNumber_r;
		pChannel^.H[stTechnoAttributeData.nFunctionNumber_r].nPrgLineNumber_r	:= stTechnoAttributeData.nPrgLineNumber_r;
		pChannel^.H[stTechnoAttributeData.nFunctionNumber_r].nFunctionNumber_r	:= stTechnoAttributeData.nFunctionNumber_r;
		pChannel^.H[stTechnoAttributeData.nFunctionNumber_r].nTime_r			:= stTechnoAttributeData.nTime_r;		
		pChannel^.H[stTechnoAttributeData.nFunctionNumber_r].bRes 				:= TRUE;	(* set acknowledge *)
		pChannel^.actH_r := CONCAT('H', UDINT_TO_STRING(stTechnoAttributeData.nFunctionNumber_r));
	ELSE
		IF NOT pChannel^.H[stTechnoAttributeData.nFunctionNumber_r].bState_rw THEN				(* wait for quit *)
			pChannel^.H[stTechnoAttributeData.nFunctionNumber_r].bRes 			:= FALSE;	(* quit the ack *)
			pChannel^.H[stTechnoAttributeData.nFunctionNumber_r].nArgument_r	:= 0;		(* reset the argument *)
			pChannel^.H[stTechnoAttributeData.nFunctionNumber_r].nBlockNumber_r		:= 0;
			pChannel^.H[stTechnoAttributeData.nFunctionNumber_r].nPrgLineNumber_r	:= 0;
			pChannel^.H[stTechnoAttributeData.nFunctionNumber_r].nFunctionNumber_r	:= 0;
			pChannel^.h[stTechnoAttributeData.nFunctionNumber_r].nTime_r			:= 0;
			pChannel^.actH_r := '';					
			bBusy 							:= FALSE;	(* quit *)
		END_IF
	END_IF
END_IF

END_FUNCTION_BLOCK

// CNC/3 Control/FB_Diag
FUNCTION_BLOCK FB_Diag
VAR_OUTPUT
	Alarm: BOOL;
	Vorwarn: BOOL;
	Meld: BOOL;
END_VAR

Alarm := TRUE;
Vorwarn := TRUE;
Meld := TRUE;

END_FUNCTION_BLOCK

// CNC/3 Control/HLI3_ChannelSetSuspendAxisOutput
FUNCTION HLI3_ChannelSetSuspendAxisOutput : BOOL
VAR_INPUT
	/// Number of channel 
	nChanIdx: INT;
	bSuspendAxis: BOOL;
END_VAR

(* ========================================================= *)
(*    FUN: HLI_ChannelSuspendAxisOutput                      *)
(* --------------------------------------------------------- *)
(*   Desc:                                                   *)
(* Author: MK , MiB                                          *)
(*   Date: 20.11.2012                                        *)
(*   Rev.: 1.1                                               *)
(* ========================================================= *)
HLI3_ChannelSetSuspendAxisOutput := TRUE;
IF NOT HLI3_CheckChannelValid(nChannel := nChanIdx) THEN
	RETURN;
END_IF
gpCh[nChanIdx]^.bahn_mc_control.suspend_axis_output.command_w := bSuspendAxis;
HLI3_ChannelSetSuspendAxisOutput := TRUE;

END_FUNCTION

// CNC/3 Control/HLI3_GetActualAxisPos
FUNCTION HLI3_GetActualAxisPos : LREAL
VAR_INPUT
	///Achs ID
	nHliAxisIdx: INT;
END_VAR
VAR
	HLI_GetActualAxisPos: DINT;
END_VAR



IF NOT (HLI3_CheckAxisValid(nHliAxisIdx := nHliAxisIdx)) THEN
	HLI3_GetActualAxisPos := -1;
	RETURN;
END_IF

HLI3_GetActualAxisPos:=  gpAx[nHliAxisIdx]^.lr_state.current_position_acs_r;

END_FUNCTION

// CNC/3 Control/HLI3_GetAxisReferenceState
FUNCTION HLI3_GetAxisReferenceState : BOOL
VAR_INPUT
	nHliAxisIdx: INT;
END_VAR


IF NOT HLI3_CheckAxisValid(nHliAxisIdx := nHliAxisIdx) THEN
	HLI3_GetAxisReferenceState := FALSE;
	RETURN;
END_IF

HLI3_GetAxisReferenceState:= gpAx[nHliAxisIdx]^.lr_state.homing_done_r;

END_FUNCTION

// CNC/3 Control/HLI3_GetAxisScaling
FUNCTION_BLOCK HLI3_GetAxisScaling
VAR_INPUT
	bExec:		BOOL;	// riding edge to start read
	nHliAxisIdx: INT;	
END_VAR
VAR_OUTPUT
	Scaling	:	LREAL;	// scalingfactor inc/0.1µm
	bBusy: 		BOOL;
	bError: 	BOOL;
	nErrorID: 	UDINT;
END_VAR
VAR
	fbAdsRead: ADSREAD;
END_VAR

(* ========================================================= *)
(*    FUN: HLI3_GetAxisScaling	                   		 	*)
(* --------------------------------------------------------- *)
(*   Desc: Gets the scaling factor of an axis   			 *)
(*															 *)
(* Return: Scaling in INC/0.1µm							 	*)
(* Author: MiB                                               *)
(* Date: 29.08.2019                                        *)
(* Rev.: 1.0                                               *)
(* ========================================================= *)



IF NOT (HLI3_CheckAxisValid(nHliAxisIdx := nHliAxisIdx)) THEN
	Scaling := 0.0;
	bError := TRUE;
	nErrorId := 1000;  // wrong HLI index
	RETURN;
END_IF


fbAdsRead(
	NETID:= '' , 
	PORT:= 551, 
	IDXGRP:= 16#23300 , 
	IDXOFFS:= 16#10000 * (nHliAxisIdx+1) + 16#1 , 
	LEN:= SIZEOF(Scaling) , 
	DESTADDR:= ADR(Scaling),
	READ:= bExec, 
	TMOUT:= , 
	BUSY=> bBusy, 
	ERR=> bError, 
	ERRID=> nErrorId );

END_FUNCTION_BLOCK

// CNC/3 Control/HLI3_GetChannelActiveG
FUNCTION_BLOCK HLI3_GetChannelActiveG
VAR_INPUT
	bExec:	   BOOL;			// riding edge to start read
	nChanIdx: INT;    			// zero based channel index	
END_VAR
VAR_OUTPUT
	ActiveG : ARRAY[0..39] OF INT;
	bBusy: BOOL;
	bError: BOOL;
	nErrorID: UDINT;
END_VAR
VAR
	fbAdsRead: ADSREAD;
END_VAR

(* ========================================================= *)
(*    FUN: HLI3_GetChannelActiveG                   		 *)
(* --------------------------------------------------------- *)
(*   Desc: Gets the channel specific active G functions      *)
(*															 *)
(* Return: Array[0..39] filled with the G information (<> -1)*)
(* Author: MiB                                               *)
(*   Date: 12.01.2016                                        *)
(*   Rev.: 1.0                                               *)
(* ========================================================= *)

fbAdsRead(
	NETID:= '' , 
	PORT:= 553, 
	IDXGRP:= 16#20100 + INT_TO_UDINT(nChanIdx) + 1, 
	IDXOFFS:= 16#3C , 
	LEN:= SIZEOF(ActiveG) , 
	DESTADDR:= ADR(ActiveG),
	READ:= bExec, 
	TMOUT:= , 
	BUSY=> bBusy, 
	ERR=> bError, 
	ERRID=> nErrorId );

END_FUNCTION_BLOCK

// CNC/3 Control/HLI3_GetChannelMessage
FUNCTION_BLOCK HLI3_GetChannelMessage
VAR_INPUT
	/// Number of channel 
	nChanIdx: INT;
	bExecute: BOOL := FALSE;
	bShowDlg: BOOL := FALSE;
END_VAR
VAR_OUTPUT
	strToPLC: STRING(HLI_MSG_CONTENT_STRL) := '';
	iMsgType: DWORD := 0;
END_VAR
VAR
	pChannel: POINTER TO HIGH_LEVEL_INTERFACE_CH;
	pMsgCU: POINTER TO MC_CONTROL_MSG_UNIT;
	pMsgToPLC: POINTER TO STRING(HLI_MSG_CONTENT_STRL);
END_VAR

(* ========================================================= *)
(*     FB: HLI_GetChannelMessage                             *)
(* --------------------------------------------------------- *)
(*   Desc: Get message from the CNC                          *)
(*   Author: MK, MiB                                         *)
(*   Date: 20.11.2012                                        *)
(*   Last:                                                   *)
(*   Rev.: 1.01                                              *)
(* ========================================================= *)

IF NOT HLI3_CheckChannelValid(nChannel := nChanIdx) THEN
	RETURN;
END_IF


(* Get pointer to data of a specific channel at the HLI *)
pChannel := gpCh[nChanIdx];

(* Control unit at the HLI that handles channel specific messages *)
pMsgCU := ADR(pChannel^.msg_mc_control);

IF bExecute = TRUE THEN
	(* Is the complete message in the control unit? *)
	IF pMsgCU^.request_semaphor_rw = TRUE
	THEN
		(* Pointer to content of the message sent to the PLC *)
		pMsgToPLC := ADR(pMsgCU^.request_r.inhalt);

		(* Get the message from the control unit *)
		strToPLC := pMsgToPLC^;

   	    CNCSystem.Channel[nChanIdx].Message := strToPLC;

		(* Get the message type *)
		iMsgType := pMsgCU^.request_r.typ;

		(* Pop up dialog with the message send to the PLC *)
		IF bShowDlg THEN
			ADSLOGSTR( msgCtrlMask := ADSLOG_MSGTYPE_MSGBOX OR ADSLOG_MSGTYPE_LOG,
			           msgFmtStr   := 'Message sent to PLC via HLI:%s',
			           strArg      := strToPLC);
		END_IF

		(* Acknowledge that you got the message *)
		pChannel^.msg_mc_control.request_semaphor_rw  := FALSE;
	END_IF;
END_IF;

END_FUNCTION_BLOCK

// CNC/3 Control/HLI3_GetFeedholdState
FUNCTION HLI3_GetFeedholdState : BOOL
VAR_INPUT
	/// Number of channel 
	nChanIdx: INT;
END_VAR


IF NOT HLI3_CheckChannelValid(nChannel := nChanIdx) THEN
	RETURN;
END_IF
HLI3_GetFeedholdState:=gpCh[nChanIdx]^.bahn_mc_control.feedhold.state_r;

END_FUNCTION

// CNC/3 Control/HLI3_GetIpoState
FUNCTION HLI3_GetIpoState : BOOL
VAR_INPUT
	nChanIdx: INT;
END_VAR



IF NOT HLI3_CheckChannelValid(nChannel := nChanIdx) THEN
	RETURN;
END_IF

HLI3_GetIpoState:=gpCh[nChanIdx]^.bahn_state.interpolation_active_r;

END_FUNCTION

// CNC/3 Control/HLI3_SetAxisGantryOn
FUNCTION HLI3_SetAxisGantryOn : BOOL
VAR_INPUT
	nHliAxisIdx: INT;
	bEnable: BOOL;
END_VAR

(****************************************************************************************)
(* POU:		HLI_SetAxisGantryOn                      									*)
(* Type:	Function																	*)
(* Author: 	HR																			*)
(* Date: 	11/01/24																	*)
(* Rev.: 	1.0																			*)
(* ------------------------------------------------------------------------------------ *)
(* Desc:	Enables the axis specific control unit for driving out the gantry			*)
(*			difference. The actual movement is triggered by the input 'bEnable'.		*)
(*			The current axis has to be a gantry slave. That means:						*)
(*				+ It is not attached to a channel										*)
(*				+ kenngr.achs_mode		0x2000n		(where n specifies the axis type)	*)
(*				+ kenngr.gantry_ax_nr	1			(e. g. axis no. of gantry master)	*)
(*				+ kenngr.gantry_offset  10000		(e. g. difference to be driven out)	*)
(*				+ kenngr.gantry_vb_korr	20000		(e. g. velocity for driving out)	*)
(****************************************************************************************)

(* Check specified logical axis no first *)
IF NOT HLI3_CheckAxisValid(nHliAxisIdx := nHliAxisIdx) THEN
	HLI3_SetAxisGantryOn := FALSE;
	RETURN;
END_IF

gpAx[nHliAxisIdx]^.lr_mc_control.gantry_on.enable_w	:= TRUE;
gpAx[nHliAxisIdx]^.lr_mc_control.gantry_on.command_w	:= bEnable;
HLI3_SetAxisGantryOn	:= TRUE;

END_FUNCTION

// CNC/3 Control/HLI3_SetAxisReferencePosition
FUNCTION HLI3_SetAxisReferencePosition : BOOL
VAR_INPUT
	bSetRefpos: BOOL;
	nHliAxisIdx: INT;
END_VAR

(* ========================================================= *)
(*    FUN: HLI_SetAxisReferenceposition                      *)
(* --------------------------------------------------------- *)
(*   Desc:                                                   *)
(* Author: HR                                                *)
(*   Date: 09.11.2010                                        *)
(*   Rev.: 1.0                                               *)
(* ========================================================= *)
HLI3_SetAxisReferencePosition := FALSE;

IF NOT HLI3_CheckAxisValid(nHliAxisIdx := nHliAxisIdx) THEN	
	RETURN;
END_IF

